   // ---------- 网络 18 ----------
   // 标题：**********************钻孔结束，枪退出速度给定*****************************************
   // 含义：条件 ((((((#DownDrillStep.S20 AND NOT (#DownDrillStep.S22)) AND ("DB720_KuKa_MainCtrl".CmdOut.gi_ToolTypeNo = 2))) AND #DownDrillStep.StopDrill_Ack) AND NOT ("DB1900_Communication_PC".Para.ProduceMode3)) AND ("DB1900_Communication_PC".Para.DrillWidth = 22.0)) 成立时，将 20 传送到 "DB1080_Component".Robot.CTRL_IN.RobotSpeed
   IF ((((((#DownDrillStep.S20 AND NOT (#DownDrillStep.S22)) AND ("DB720_KuKa_MainCtrl".CmdOut.gi_ToolTypeNo = 2))) AND #DownDrillStep.StopDrill_Ack) AND NOT ("DB1900_Communication_PC".Para.ProduceMode3)) AND ("DB1900_Communication_PC".Para.DrillWidth = 22.0)) THEN
       "DB1080_Component".Robot.CTRL_IN.RobotSpeed := 20;
   END_IF;
   // 含义：条件 ((((((#DownDrillStep.S20 AND NOT (#DownDrillStep.S22)) AND ("DB720_KuKa_MainCtrl".CmdOut.gi_ToolTypeNo = 2))) AND #DownDrillStep.StopDrill_Ack) AND NOT ("DB1900_Communication_PC".Para.ProduceMode3)) AND ("DB1900_Communication_PC".Para.DrillWidth = 25.0)) 成立时，将 25 传送到 "DB1080_Component".Robot.CTRL_IN.RobotSpeed
   IF ((((((#DownDrillStep.S20 AND NOT (#DownDrillStep.S22)) AND ("DB720_KuKa_MainCtrl".CmdOut.gi_ToolTypeNo = 2))) AND #DownDrillStep.StopDrill_Ack) AND NOT ("DB1900_Communication_PC".Para.ProduceMode3)) AND ("DB1900_Communication_PC".Para.DrillWidth = 25.0)) THEN
       "DB1080_Component".Robot.CTRL_IN.RobotSpeed := 25;
   END_IF;
   // 含义：条件 ((((((#DownDrillStep.S20 AND NOT (#DownDrillStep.S22)) AND ("DB720_KuKa_MainCtrl".CmdOut.gi_ToolTypeNo = 2))) AND #DownDrillStep.StopDrill_Ack) AND NOT ("DB1900_Communication_PC".Para.ProduceMode3)) AND ("DB1900_Communication_PC".Para.DrillWidth > 25.0)) 成立时，将 30 传送到 "DB1080_Component".Robot.CTRL_IN.RobotSpeed
   IF ((((((#DownDrillStep.S20 AND NOT (#DownDrillStep.S22)) AND ("DB720_KuKa_MainCtrl".CmdOut.gi_ToolTypeNo = 2))) AND #DownDrillStep.StopDrill_Ack) AND NOT ("DB1900_Communication_PC".Para.ProduceMode3)) AND ("DB1900_Communication_PC".Para.DrillWidth > 25.0)) THEN
       "DB1080_Component".Robot.CTRL_IN.RobotSpeed := 30;
   END_IF;
   // 含义：条件 ((((#DownDrillStep.S20 AND NOT (#DownDrillStep.S22)) AND ("DB720_KuKa_MainCtrl".CmdOut.gi_ToolTypeNo = 2))) AND #DownDrillStep.StopDrill_Ack) AND "DB1900_Communication_PC".Para.ProduceMode3 成立时，将 50 传送到 "DB1080_Component".Robot.CTRL_IN.RobotSpeed
   IF ((((#DownDrillStep.S20 AND NOT (#DownDrillStep.S22)) AND ("DB720_KuKa_MainCtrl".CmdOut.gi_ToolTypeNo = 2))) AND #DownDrillStep.StopDrill_Ack) AND "DB1900_Communication_PC".Para.ProduceMode3 THEN
       "DB1080_Component".Robot.CTRL_IN.RobotSpeed := 50;
   END_IF;
   // 含义：条件 ((((((#DownDrillStep.S20 AND NOT (#DownDrillStep.S22)) AND ("DB720_KuKa_MainCtrl".CmdOut.gi_ToolTypeNo = 13))) AND #Aux.StartDrill) AND NOT (#DownDrillStep.StopDrill_Ack)) AND ("DB1900_Communication_PC".Recv.Current_2 > 12.0)) 成立时，将 1 传送到 "DB1080_Component".Robot.CTRL_IN.RobotSpeed
   IF ((((((#DownDrillStep.S20 AND NOT (#DownDrillStep.S22)) AND ("DB720_KuKa_MainCtrl".CmdOut.gi_ToolTypeNo = 13))) AND #Aux.StartDrill) AND NOT (#DownDrillStep.StopDrill_Ack)) AND ("DB1900_Communication_PC".Recv.Current_2 > 12.0)) THEN
       "DB1080_Component".Robot.CTRL_IN.RobotSpeed := 1;
   END_IF;
   // 含义：条件 ((((((#DownDrillStep.S20 AND NOT (#DownDrillStep.S22)) AND ("DB720_KuKa_MainCtrl".CmdOut.gi_ToolTypeNo = 13))) AND #Aux.StartDrill) AND #DownDrillStep.StopDrill_Ack) AND ("DB1900_Communication_PC".Recv.Current_2 < 12.0)) 成立时，将 30 传送到 "DB1080_Component".Robot.CTRL_IN.RobotSpeed
   IF ((((((#DownDrillStep.S20 AND NOT (#DownDrillStep.S22)) AND ("DB720_KuKa_MainCtrl".CmdOut.gi_ToolTypeNo = 13))) AND #Aux.StartDrill) AND #DownDrillStep.StopDrill_Ack) AND ("DB1900_Communication_PC".Recv.Current_2 < 12.0)) THEN
       "DB1080_Component".Robot.CTRL_IN.RobotSpeed := 30;
   END_IF;
   // 含义：条件 ((((((#DownDrillStep.S20 AND NOT (#DownDrillStep.S22)) AND ("DB720_KuKa_MainCtrl".CmdOut.gi_ToolTypeNo = 13))) AND #Aux.StartDrill) AND #DownDrillStep.StopDrill_Ack) AND ("DB1900_Communication_PC".Recv.Current_2 >= 12.0)) 成立时，将 10 传送到 "DB1080_Component".Robot.CTRL_IN.RobotSpeed
   IF ((((((#DownDrillStep.S20 AND NOT (#DownDrillStep.S22)) AND ("DB720_KuKa_MainCtrl".CmdOut.gi_ToolTypeNo = 13))) AND #Aux.StartDrill) AND #DownDrillStep.StopDrill_Ack) AND ("DB1900_Communication_PC".Recv.Current_2 >= 12.0)) THEN
       "DB1080_Component".Robot.CTRL_IN.RobotSpeed := 10;
   END_IF;

   // ---------- 网络 19 ----------
   // 标题：****************故障计数（包含钻超时，低电流，打孔深度超限）**************************
   // 含义：调用计数器实例 "Timer_DownChiselEnd".TON（上升沿计数，当前值写入 CV）
   "Timer_DownChiselEnd".TON(IN := ((((#DownDrillStep.S20 AND NOT (#DownDrillStep.S22)) AND "DB1900_Communication_PC".Para.ProduceMode3) AND "DB720_KuKa_MainCtrl".StatusIn.do_DrilEnd_Pos) AND ("DB1900_Communication_PC".Recv.Current_2 < "DB1900_Communication_PC".Para.CurrentMinLimit)),
                             PT := T#3s);
   // 含义：条件 "Timer_DownChiselEnd".Q 成立时，将 TRUE 传送到 "DB1060_AutoStep".DownDrillAutoStep.DownDrillStep.ChiselEndPos
   IF "Timer_DownChiselEnd".Q THEN
       "DB1060_AutoStep".DownDrillAutoStep.DownDrillStep.ChiselEndPos := TRUE;
   END_IF;
   // 含义：条件 "Timer_DownChiselEnd".Q 成立时，将 ("DB1042_Timer".DCLowTimeOutTimes + 1) 传送到 "DB1042_Timer".DCLowTimeOutTimes
   IF "Timer_DownChiselEnd".Q THEN
       "DB1042_Timer".DCLowTimeOutTimes := ("DB1042_Timer".DCLowTimeOutTimes + 1);
   END_IF;
   // 含义：条件 (((((#DownDrillStep.S20 AND NOT (#DownDrillStep.S22)) AND "DB1900_Communication_PC".Para.ProduceMode3) AND ("DB1900_Communication_PC".Recv.Current_2 > "DB1900_Communication_PC".Para.CurrentMinLimit))) AND ("DB1900_Communication_PC".Recv.Current_2 < "DB1900_Communication_PC".Para.CurrentMaxLimit)) 成立时，将 0 传送到 "DB1042_Timer".DCLowTimeOutTimes
   IF (((((#DownDrillStep.S20 AND NOT (#DownDrillStep.S22)) AND "DB1900_Communication_PC".Para.ProduceMode3) AND ("DB1900_Communication_PC".Recv.Current_2 > "DB1900_Communication_PC".Para.CurrentMinLimit))) AND ("DB1900_Communication_PC".Recv.Current_2 < "DB1900_Communication_PC".Para.CurrentMaxLimit)) THEN
       "DB1042_Timer".DCLowTimeOutTimes := 0;
   END_IF;
   // 含义：条件 ((((#DownDrillStep.S20 AND NOT (#DownDrillStep.S22)) AND "DB1900_Communication_PC".Para.ProduceMode3) AND "DB1042_Timer".DDrillEndTime.Q) OR (((#DownDrillStep.S20 AND NOT (#DownDrillStep.S22)) AND "DB1900_Communication_PC".Para.ProduceMode3) AND #Aux.DDrillTime.Q) OR (((#DownDrillStep.S20 AND NOT (#DownDrillStep.S22)) AND "DB1900_Communication_PC".Para.ProduceMode3) AND "DB1042_Timer".CurrentLowTimeOut.Q) OR (((#DownDrillStep.S20 AND NOT (#DownDrillStep.S22)) AND "DB1900_Communication_PC".Para.ProduceMode3) AND "DB1042_Timer".CurrentHighTimeOut.Q) OR (((#DownDrillStep.S20 AND NOT (#DownDrillStep.S22)) AND "DB1900_Communication_PC".Para.ProduceMode3) AND "DB1060_AutoStep".DownDrillAutoStep.DownDrillStep.ChiselEndPos) OR ((((#DownDrillStep.S20 AND NOT (#DownDrillStep.S22)) AND "DB1900_Communication_PC".Para.ProduceMode3) AND ("DB1900_Communication_PC".Send.ScrLen >= "DB1900_Communication_PC".Para.DrillDepth)))) AND NOT ("DB720_KuKa_MainCtrl".StatusIn.do_ChiselCylinderExt) 成立时，将 0.0 传送到 "DB1080_Component".Aux.Pressure
   IF ((((#DownDrillStep.S20 AND NOT (#DownDrillStep.S22)) AND "DB1900_Communication_PC".Para.ProduceMode3) AND "DB1042_Timer".DDrillEndTime.Q) OR (((#DownDrillStep.S20 AND NOT (#DownDrillStep.S22)) AND "DB1900_Communication_PC".Para.ProduceMode3) AND #Aux.DDrillTime.Q) OR (((#DownDrillStep.S20 AND NOT (#DownDrillStep.S22)) AND "DB1900_Communication_PC".Para.ProduceMode3) AND "DB1042_Timer".CurrentLowTimeOut.Q) OR (((#DownDrillStep.S20 AND NOT (#DownDrillStep.S22)) AND "DB1900_Communication_PC".Para.ProduceMode3) AND "DB1042_Timer".CurrentHighTimeOut.Q) OR (((#DownDrillStep.S20 AND NOT (#DownDrillStep.S22)) AND "DB1900_Communication_PC".Para.ProduceMode3) AND "DB1060_AutoStep".DownDrillAutoStep.DownDrillStep.ChiselEndPos) OR ((((#DownDrillStep.S20 AND NOT (#DownDrillStep.S22)) AND "DB1900_Communication_PC".Para.ProduceMode3) AND ("DB1900_Communication_PC".Send.ScrLen >= "DB1900_Communication_PC".Para.DrillDepth)))) AND NOT ("DB720_KuKa_MainCtrl".StatusIn.do_ChiselCylinderExt) THEN
       "DB1080_Component".Aux.Pressure := 0.0;
   END_IF;
   // 含义：条件 ((((#DownDrillStep.S20 AND NOT (#DownDrillStep.S22)) AND "DB1900_Communication_PC".Para.ProduceMode3) AND "DB1042_Timer".DDrillEndTime.Q) OR (((#DownDrillStep.S20 AND NOT (#DownDrillStep.S22)) AND "DB1900_Communication_PC".Para.ProduceMode3) AND #Aux.DDrillTime.Q) OR (((#DownDrillStep.S20 AND NOT (#DownDrillStep.S22)) AND "DB1900_Communication_PC".Para.ProduceMode3) AND "DB1042_Timer".CurrentLowTimeOut.Q) OR (((#DownDrillStep.S20 AND NOT (#DownDrillStep.S22)) AND "DB1900_Communication_PC".Para.ProduceMode3) AND "DB1042_Timer".CurrentHighTimeOut.Q) OR (((#DownDrillStep.S20 AND NOT (#DownDrillStep.S22)) AND "DB1900_Communication_PC".Para.ProduceMode3) AND "DB1060_AutoStep".DownDrillAutoStep.DownDrillStep.ChiselEndPos) OR ((((#DownDrillStep.S20 AND NOT (#DownDrillStep.S22)) AND "DB1900_Communication_PC".Para.ProduceMode3) AND ("DB1900_Communication_PC".Send.ScrLen >= "DB1900_Communication_PC".Para.DrillDepth)))) AND NOT ("DB720_KuKa_MainCtrl".CmdOut.di_ChiselRobotRet) 成立时，将 TRUE 传送到 "DB1081_ValveCall".ST01.Z02.RetAuto
   IF ((((#DownDrillStep.S20 AND NOT (#DownDrillStep.S22)) AND "DB1900_Communication_PC".Para.ProduceMode3) AND "DB1042_Timer".DDrillEndTime.Q) OR (((#DownDrillStep.S20 AND NOT (#DownDrillStep.S22)) AND "DB1900_Communication_PC".Para.ProduceMode3) AND #Aux.DDrillTime.Q) OR (((#DownDrillStep.S20 AND NOT (#DownDrillStep.S22)) AND "DB1900_Communication_PC".Para.ProduceMode3) AND "DB1042_Timer".CurrentLowTimeOut.Q) OR (((#DownDrillStep.S20 AND NOT (#DownDrillStep.S22)) AND "DB1900_Communication_PC".Para.ProduceMode3) AND "DB1042_Timer".CurrentHighTimeOut.Q) OR (((#DownDrillStep.S20 AND NOT (#DownDrillStep.S22)) AND "DB1900_Communication_PC".Para.ProduceMode3) AND "DB1060_AutoStep".DownDrillAutoStep.DownDrillStep.ChiselEndPos) OR ((((#DownDrillStep.S20 AND NOT (#DownDrillStep.S22)) AND "DB1900_Communication_PC".Para.ProduceMode3) AND ("DB1900_Communication_PC".Send.ScrLen >= "DB1900_Communication_PC".Para.DrillDepth)))) AND NOT ("DB720_KuKa_MainCtrl".CmdOut.di_ChiselRobotRet) THEN
       "DB1081_ValveCall".ST01.Z02.RetAuto := TRUE;
   END_IF;
   // 含义：条件 ((((#DownDrillStep.S20 AND NOT (#DownDrillStep.S22)) AND "DB1900_Communication_PC".Para.ProduceMode3) AND "DB1042_Timer".DDrillEndTime.Q) OR (((#DownDrillStep.S20 AND NOT (#DownDrillStep.S22)) AND "DB1900_Communication_PC".Para.ProduceMode3) AND #Aux.DDrillTime.Q) OR (((#DownDrillStep.S20 AND NOT (#DownDrillStep.S22)) AND "DB1900_Communication_PC".Para.ProduceMode3) AND "DB1042_Timer".CurrentLowTimeOut.Q) OR (((#DownDrillStep.S20 AND NOT (#DownDrillStep.S22)) AND "DB1900_Communication_PC".Para.ProduceMode3) AND "DB1042_Timer".CurrentHighTimeOut.Q) OR (((#DownDrillStep.S20 AND NOT (#DownDrillStep.S22)) AND "DB1900_Communication_PC".Para.ProduceMode3) AND "DB1060_AutoStep".DownDrillAutoStep.DownDrillStep.ChiselEndPos) OR ((((#DownDrillStep.S20 AND NOT (#DownDrillStep.S22)) AND "DB1900_Communication_PC".Para.ProduceMode3) AND ("DB1900_Communication_PC".Send.ScrLen >= "DB1900_Communication_PC".Para.DrillDepth)))) AND "DB720_KuKa_MainCtrl".StatusIn.do_ChiselCylinderExt 成立时，将 FALSE 传送到 "DB1081_ValveCall".ST01.Z02.RetAuto
   IF ((((#DownDrillStep.S20 AND NOT (#DownDrillStep.S22)) AND "DB1900_Communication_PC".Para.ProduceMode3) AND "DB1042_Timer".DDrillEndTime.Q) OR (((#DownDrillStep.S20 AND NOT (#DownDrillStep.S22)) AND "DB1900_Communication_PC".Para.ProduceMode3) AND #Aux.DDrillTime.Q) OR (((#DownDrillStep.S20 AND NOT (#DownDrillStep.S22)) AND "DB1900_Communication_PC".Para.ProduceMode3) AND "DB1042_Timer".CurrentLowTimeOut.Q) OR (((#DownDrillStep.S20 AND NOT (#DownDrillStep.S22)) AND "DB1900_Communication_PC".Para.ProduceMode3) AND "DB1042_Timer".CurrentHighTimeOut.Q) OR (((#DownDrillStep.S20 AND NOT (#DownDrillStep.S22)) AND "DB1900_Communication_PC".Para.ProduceMode3) AND "DB1060_AutoStep".DownDrillAutoStep.DownDrillStep.ChiselEndPos) OR ((((#DownDrillStep.S20 AND NOT (#DownDrillStep.S22)) AND "DB1900_Communication_PC".Para.ProduceMode3) AND ("DB1900_Communication_PC".Send.ScrLen >= "DB1900_Communication_PC".Para.DrillDepth)))) AND "DB720_KuKa_MainCtrl".StatusIn.do_ChiselCylinderExt THEN
       "DB1081_ValveCall".ST01.Z02.RetAuto := FALSE;
   END_IF;
   // 含义：条件 ((((#DownDrillStep.S20 AND NOT (#DownDrillStep.S22)) AND "DB1900_Communication_PC".Para.ProduceMode3) AND "DB1042_Timer".DDrillEndTime.Q) OR (((#DownDrillStep.S20 AND NOT (#DownDrillStep.S22)) AND "DB1900_Communication_PC".Para.ProduceMode3) AND #Aux.DDrillTime.Q) OR (((#DownDrillStep.S20 AND NOT (#DownDrillStep.S22)) AND "DB1900_Communication_PC".Para.ProduceMode3) AND "DB1042_Timer".CurrentLowTimeOut.Q) OR (((#DownDrillStep.S20 AND NOT (#DownDrillStep.S22)) AND "DB1900_Communication_PC".Para.ProduceMode3) AND "DB1042_Timer".CurrentHighTimeOut.Q) OR (((#DownDrillStep.S20 AND NOT (#DownDrillStep.S22)) AND "DB1900_Communication_PC".Para.ProduceMode3) AND "DB1060_AutoStep".DownDrillAutoStep.DownDrillStep.ChiselEndPos) OR ((((#DownDrillStep.S20 AND NOT (#DownDrillStep.S22)) AND "DB1900_Communication_PC".Para.ProduceMode3) AND ("DB1900_Communication_PC".Send.ScrLen >= "DB1900_Communication_PC".Para.DrillDepth)))) AND "DB720_KuKa_MainCtrl".StatusIn.do_ReqStopDril 成立时，将 FALSE 传送到 "DB720_KuKa_MainCtrl".CmdOut.di_ChiselCylinderRet
   IF ((((#DownDrillStep.S20 AND NOT (#DownDrillStep.S22)) AND "DB1900_Communication_PC".Para.ProduceMode3) AND "DB1042_Timer".DDrillEndTime.Q) OR (((#DownDrillStep.S20 AND NOT (#DownDrillStep.S22)) AND "DB1900_Communication_PC".Para.ProduceMode3) AND #Aux.DDrillTime.Q) OR (((#DownDrillStep.S20 AND NOT (#DownDrillStep.S22)) AND "DB1900_Communication_PC".Para.ProduceMode3) AND "DB1042_Timer".CurrentLowTimeOut.Q) OR (((#DownDrillStep.S20 AND NOT (#DownDrillStep.S22)) AND "DB1900_Communication_PC".Para.ProduceMode3) AND "DB1042_Timer".CurrentHighTimeOut.Q) OR (((#DownDrillStep.S20 AND NOT (#DownDrillStep.S22)) AND "DB1900_Communication_PC".Para.ProduceMode3) AND "DB1060_AutoStep".DownDrillAutoStep.DownDrillStep.ChiselEndPos) OR ((((#DownDrillStep.S20 AND NOT (#DownDrillStep.S22)) AND "DB1900_Communication_PC".Para.ProduceMode3) AND ("DB1900_Communication_PC".Send.ScrLen >= "DB1900_Communication_PC".Para.DrillDepth)))) AND "DB720_KuKa_MainCtrl".StatusIn.do_ReqStopDril THEN
       "DB720_KuKa_MainCtrl".CmdOut.di_ChiselCylinderRet := FALSE;
   END_IF;
   // 含义：条件 ((((#DownDrillStep.S20 AND NOT (#DownDrillStep.S22)) AND "DB1900_Communication_PC".Para.ProduceMode3) AND "DB1042_Timer".DDrillEndTime.Q) OR (((#DownDrillStep.S20 AND NOT (#DownDrillStep.S22)) AND "DB1900_Communication_PC".Para.ProduceMode3) AND #Aux.DDrillTime.Q) OR (((#DownDrillStep.S20 AND NOT (#DownDrillStep.S22)) AND "DB1900_Communication_PC".Para.ProduceMode3) AND "DB1042_Timer".CurrentLowTimeOut.Q) OR (((#DownDrillStep.S20 AND NOT (#DownDrillStep.S22)) AND "DB1900_Communication_PC".Para.ProduceMode3) AND "DB1042_Timer".CurrentHighTimeOut.Q) OR (((#DownDrillStep.S20 AND NOT (#DownDrillStep.S22)) AND "DB1900_Communication_PC".Para.ProduceMode3) AND "DB1060_AutoStep".DownDrillAutoStep.DownDrillStep.ChiselEndPos) OR ((((#DownDrillStep.S20 AND NOT (#DownDrillStep.S22)) AND "DB1900_Communication_PC".Para.ProduceMode3) AND ("DB1900_Communication_PC".Send.ScrLen >= "DB1900_Communication_PC".Para.DrillDepth)))) AND "DB720_KuKa_MainCtrl".StatusIn.do_ReqStopDril 成立时，将 FALSE 传送到 "DB720_KuKa_MainCtrl".CmdOut.di_ChiselRobotRet
   IF ((((#DownDrillStep.S20 AND NOT (#DownDrillStep.S22)) AND "DB1900_Communication_PC".Para.ProduceMode3) AND "DB1042_Timer".DDrillEndTime.Q) OR (((#DownDrillStep.S20 AND NOT (#DownDrillStep.S22)) AND "DB1900_Communication_PC".Para.ProduceMode3) AND #Aux.DDrillTime.Q) OR (((#DownDrillStep.S20 AND NOT (#DownDrillStep.S22)) AND "DB1900_Communication_PC".Para.ProduceMode3) AND "DB1042_Timer".CurrentLowTimeOut.Q) OR (((#DownDrillStep.S20 AND NOT (#DownDrillStep.S22)) AND "DB1900_Communication_PC".Para.ProduceMode3) AND "DB1042_Timer".CurrentHighTimeOut.Q) OR (((#DownDrillStep.S20 AND NOT (#DownDrillStep.S22)) AND "DB1900_Communication_PC".Para.ProduceMode3) AND "DB1060_AutoStep".DownDrillAutoStep.DownDrillStep.ChiselEndPos) OR ((((#DownDrillStep.S20 AND NOT (#DownDrillStep.S22)) AND "DB1900_Communication_PC".Para.ProduceMode3) AND ("DB1900_Communication_PC".Send.ScrLen >= "DB1900_Communication_PC".Para.DrillDepth)))) AND "DB720_KuKa_MainCtrl".StatusIn.do_ReqStopDril THEN
       "DB720_KuKa_MainCtrl".CmdOut.di_ChiselRobotRet := FALSE;
   END_IF;
   // 含义：条件 ((((((#DownDrillStep.S20 AND NOT (#DownDrillStep.S22)) AND "DB1900_Communication_PC".Para.ProduceMode3) AND "DB1042_Timer".DDrillEndTime.Q) OR (((#DownDrillStep.S20 AND NOT (#DownDrillStep.S22)) AND "DB1900_Communication_PC".Para.ProduceMode3) AND #Aux.DDrillTime.Q) OR (((#DownDrillStep.S20 AND NOT (#DownDrillStep.S22)) AND "DB1900_Communication_PC".Para.ProduceMode3) AND "DB1042_Timer".CurrentLowTimeOut.Q) OR (((#DownDrillStep.S20 AND NOT (#DownDrillStep.S22)) AND "DB1900_Communication_PC".Para.ProduceMode3) AND "DB1042_Timer".CurrentHighTimeOut.Q) OR (((#DownDrillStep.S20 AND NOT (#DownDrillStep.S22)) AND "DB1900_Communication_PC".Para.ProduceMode3) AND "DB1060_AutoStep".DownDrillAutoStep.DownDrillStep.ChiselEndPos) OR ((((#DownDrillStep.S20 AND NOT (#DownDrillStep.S22)) AND "DB1900_Communication_PC".Para.ProduceMode3) AND ("DB1900_Communication_PC".Send.ScrLen >= "DB1900_Communication_PC".Para.DrillDepth)))) AND "IZ02RetPos") AND ("DB1080_Component".ClinyderPos.Ctrl_Out.Cur_Val_Out >= 92.5)) 成立时，将 TRUE 传送到 "DB720_KuKa_MainCtrl".CmdOut.di_ChiselCylinderRet
   IF ((((((#DownDrillStep.S20 AND NOT (#DownDrillStep.S22)) AND "DB1900_Communication_PC".Para.ProduceMode3) AND "DB1042_Timer".DDrillEndTime.Q) OR (((#DownDrillStep.S20 AND NOT (#DownDrillStep.S22)) AND "DB1900_Communication_PC".Para.ProduceMode3) AND #Aux.DDrillTime.Q) OR (((#DownDrillStep.S20 AND NOT (#DownDrillStep.S22)) AND "DB1900_Communication_PC".Para.ProduceMode3) AND "DB1042_Timer".CurrentLowTimeOut.Q) OR (((#DownDrillStep.S20 AND NOT (#DownDrillStep.S22)) AND "DB1900_Communication_PC".Para.ProduceMode3) AND "DB1042_Timer".CurrentHighTimeOut.Q) OR (((#DownDrillStep.S20 AND NOT (#DownDrillStep.S22)) AND "DB1900_Communication_PC".Para.ProduceMode3) AND "DB1060_AutoStep".DownDrillAutoStep.DownDrillStep.ChiselEndPos) OR ((((#DownDrillStep.S20 AND NOT (#DownDrillStep.S22)) AND "DB1900_Communication_PC".Para.ProduceMode3) AND ("DB1900_Communication_PC".Send.ScrLen >= "DB1900_Communication_PC".Para.DrillDepth)))) AND "IZ02RetPos") AND ("DB1080_Component".ClinyderPos.Ctrl_Out.Cur_Val_Out >= 92.5)) THEN
       "DB720_KuKa_MainCtrl".CmdOut.di_ChiselCylinderRet := TRUE;
   END_IF;
   // 含义：条件 ((((((#DownDrillStep.S20 AND NOT (#DownDrillStep.S22)) AND "DB1900_Communication_PC".Para.ProduceMode3) AND "DB1042_Timer".DDrillEndTime.Q) OR (((#DownDrillStep.S20 AND NOT (#DownDrillStep.S22)) AND "DB1900_Communication_PC".Para.ProduceMode3) AND #Aux.DDrillTime.Q) OR (((#DownDrillStep.S20 AND NOT (#DownDrillStep.S22)) AND "DB1900_Communication_PC".Para.ProduceMode3) AND "DB1042_Timer".CurrentLowTimeOut.Q) OR (((#DownDrillStep.S20 AND NOT (#DownDrillStep.S22)) AND "DB1900_Communication_PC".Para.ProduceMode3) AND "DB1042_Timer".CurrentHighTimeOut.Q) OR (((#DownDrillStep.S20 AND NOT (#DownDrillStep.S22)) AND "DB1900_Communication_PC".Para.ProduceMode3) AND "DB1060_AutoStep".DownDrillAutoStep.DownDrillStep.ChiselEndPos) OR ((((#DownDrillStep.S20 AND NOT (#DownDrillStep.S22)) AND "DB1900_Communication_PC".Para.ProduceMode3) AND ("DB1900_Communication_PC".Send.ScrLen >= "DB1900_Communication_PC".Para.DrillDepth)))) AND "IZ02RetPos") AND ("DB1080_Component".ClinyderPos.Ctrl_Out.Cur_Val_Out >= 92.5)) 成立时，将 TRUE 传送到 "DB720_KuKa_MainCtrl".CmdOut.di_ChiselRobotRet
   IF ((((((#DownDrillStep.S20 AND NOT (#DownDrillStep.S22)) AND "DB1900_Communication_PC".Para.ProduceMode3) AND "DB1042_Timer".DDrillEndTime.Q) OR (((#DownDrillStep.S20 AND NOT (#DownDrillStep.S22)) AND "DB1900_Communication_PC".Para.ProduceMode3) AND #Aux.DDrillTime.Q) OR (((#DownDrillStep.S20 AND NOT (#DownDrillStep.S22)) AND "DB1900_Communication_PC".Para.ProduceMode3) AND "DB1042_Timer".CurrentLowTimeOut.Q) OR (((#DownDrillStep.S20 AND NOT (#DownDrillStep.S22)) AND "DB1900_Communication_PC".Para.ProduceMode3) AND "DB1042_Timer".CurrentHighTimeOut.Q) OR (((#DownDrillStep.S20 AND NOT (#DownDrillStep.S22)) AND "DB1900_Communication_PC".Para.ProduceMode3) AND "DB1060_AutoStep".DownDrillAutoStep.DownDrillStep.ChiselEndPos) OR ((((#DownDrillStep.S20 AND NOT (#DownDrillStep.S22)) AND "DB1900_Communication_PC".Para.ProduceMode3) AND ("DB1900_Communication_PC".Send.ScrLen >= "DB1900_Communication_PC".Para.DrillDepth)))) AND "IZ02RetPos") AND ("DB1080_Component".ClinyderPos.Ctrl_Out.Cur_Val_Out >= 92.5)) THEN
       "DB720_KuKa_MainCtrl".CmdOut.di_ChiselRobotRet := TRUE;
   END_IF;
   // 含义：调用计数器实例 "Timer_CylinderBack_Down".TON（上升沿计数，当前值写入 CV）
   "Timer_CylinderBack_Down".TON(IN := ((((#DownDrillStep.S20 AND NOT (#DownDrillStep.S22)) AND "DB1900_Communication_PC".Para.ProduceMode3) AND "DB1042_Timer".DDrillEndTime.Q) OR (((#DownDrillStep.S20 AND NOT (#DownDrillStep.S22)) AND "DB1900_Communication_PC".Para.ProduceMode3) AND #Aux.DDrillTime.Q) OR (((#DownDrillStep.S20 AND NOT (#DownDrillStep.S22)) AND "DB1900_Communication_PC".Para.ProduceMode3) AND "DB1042_Timer".CurrentLowTimeOut.Q) OR (((#DownDrillStep.S20 AND NOT (#DownDrillStep.S22)) AND "DB1900_Communication_PC".Para.ProduceMode3) AND "DB1042_Timer".CurrentHighTimeOut.Q) OR (((#DownDrillStep.S20 AND NOT (#DownDrillStep.S22)) AND "DB1900_Communication_PC".Para.ProduceMode3) AND "DB1060_AutoStep".DownDrillAutoStep.DownDrillStep.ChiselEndPos) OR ((((#DownDrillStep.S20 AND NOT (#DownDrillStep.S22)) AND "DB1900_Communication_PC".Para.ProduceMode3) AND ("DB1900_Communication_PC".Send.ScrLen >= "DB1900_Communication_PC".Para.DrillDepth)))) AND NOT ("IZ02RetPos"),
                                 PT := t#3s);
   // 含义：条件 "Timer_CylinderBack_Down".Q 成立时，将 TRUE 传送到 "DB720_KuKa_MainCtrl".CmdOut.di_ChiselRobotRet
   IF "Timer_CylinderBack_Down".Q THEN
       "DB720_KuKa_MainCtrl".CmdOut.di_ChiselRobotRet := TRUE;
   END_IF;
   // 含义：调用计数器实例 "Timer_RobotPry_Down".TON（上升沿计数，当前值写入 CV）
   "Timer_RobotPry_Down".TON(IN := (((((#DownDrillStep.S20 AND NOT (#DownDrillStep.S22)) AND "DB1900_Communication_PC".Para.ProduceMode3) AND "DB1042_Timer".DDrillEndTime.Q) OR (((#DownDrillStep.S20 AND NOT (#DownDrillStep.S22)) AND "DB1900_Communication_PC".Para.ProduceMode3) AND #Aux.DDrillTime.Q) OR (((#DownDrillStep.S20 AND NOT (#DownDrillStep.S22)) AND "DB1900_Communication_PC".Para.ProduceMode3) AND "DB1042_Timer".CurrentLowTimeOut.Q) OR (((#DownDrillStep.S20 AND NOT (#DownDrillStep.S22)) AND "DB1900_Communication_PC".Para.ProduceMode3) AND "DB1042_Timer".CurrentHighTimeOut.Q) OR (((#DownDrillStep.S20 AND NOT (#DownDrillStep.S22)) AND "DB1900_Communication_PC".Para.ProduceMode3) AND "DB1060_AutoStep".DownDrillAutoStep.DownDrillStep.ChiselEndPos) OR ((((#DownDrillStep.S20 AND NOT (#DownDrillStep.S22)) AND "DB1900_Communication_PC".Para.ProduceMode3) AND ("DB1900_Communication_PC".Send.ScrLen >= "DB1900_Communication_PC".Para.DrillDepth)))) AND NOT ("IZ02RetPos")) AND "DB720_KuKa_MainCtrl".StatusIn.do_RobotPry_End,
                             PT := t#3s);
   // 含义：条件 "Timer_RobotPry_Down".Q 成立时，将 FALSE 传送到 "DB720_KuKa_MainCtrl".CmdOut.di_ChiselCylinderRet
   IF "Timer_RobotPry_Down".Q THEN
       "DB720_KuKa_MainCtrl".CmdOut.di_ChiselCylinderRet := FALSE;
   END_IF;
   // 含义：条件 "Timer_RobotPry_Down".Q 成立时，将 FALSE 传送到 "DB720_KuKa_MainCtrl".CmdOut.di_ChiselRobotRet
   IF "Timer_RobotPry_Down".Q THEN
       "DB720_KuKa_MainCtrl".CmdOut.di_ChiselRobotRet := FALSE;
   END_IF;
   // 含义：条件 "Timer_RobotPry_Down".Q 成立时，将 TRUE 传送到 "DB1148_PromptBeeper".Public.DownChiselStuckErr
   IF "Timer_RobotPry_Down".Q THEN
       "DB1148_PromptBeeper".Public.DownChiselStuckErr := TRUE;
   END_IF;
   // 含义：条件 "Timer_RobotPry_Down".Q 成立时，将 TRUE 传送到 #DownDrillStep.ErrEnd
   IF "Timer_RobotPry_Down".Q THEN
       #DownDrillStep.ErrEnd := TRUE;
   END_IF;
   // 含义：条件 "Timer_RobotPry_Down".Q 成立时，将 FALSE 传送到 "DB1081_ValveCall".ST01.Z02.RetAuto
   IF "Timer_RobotPry_Down".Q THEN
       "DB1081_ValveCall".ST01.Z02.RetAuto := FALSE;
   END_IF;
   // 含义：条件 "Timer_RobotPry_Down".Q 成立时，将 TRUE 传送到 "DB1081_ValveCall".ST01.Z01.ExtAuto
   IF "Timer_RobotPry_Down".Q THEN
       "DB1081_ValveCall".ST01.Z01.ExtAuto := TRUE;
   END_IF;
   // 含义：条件 "Timer_RobotPry_Down".Q 成立时，将 FALSE 传送到 "DB1081_ValveCall".ST01.Z01.RetAuto
   IF "Timer_RobotPry_Down".Q THEN
       "DB1081_ValveCall".ST01.Z01.RetAuto := FALSE;
   END_IF;
   // 含义：条件 "Timer_RobotPry_Down".Q 成立时，将 0.1 传送到 "DB1080_Component".Aux.Pressure
   IF "Timer_RobotPry_Down".Q THEN
       "DB1080_Component".Aux.Pressure := 0.1;
   END_IF;
   // 含义：将 (((#DownDrillStep.S20 AND NOT (#DownDrillStep.S22)) AND #Aux.DDrillTime.Q) OR ((#DownDrillStep.S20 AND NOT (#DownDrillStep.S22)) AND "DB1042_Timer".CurrentLowTimeOut.Q) OR ((#DownDrillStep.S20 AND NOT (#DownDrillStep.S22)) AND "DB1042_Timer".CurrentHighTimeOut.Q) OR ((((((((#DownDrillStep.S20 AND NOT (#DownDrillStep.S22)) AND NOT ("DB1900_Communication_PC".Para.ProduceMode3)) AND ("DB1900_Communication_PC".Send.PosNo <= 2))) AND ("DB1900_Communication_PC".Para.DrillWidth <= 28.0))) AND ("DB1900_Communication_PC".Send.ScrLen >= 55.0))) OR ((((#DownDrillStep.S20 AND NOT (#DownDrillStep.S22)) AND NOT ("DB1900_Communication_PC".Para.ProduceMode3)) AND ("DB1900_Communication_PC".Send.ScrLen >= "DB1900_Communication_PC".Para.DrillDepth))) OR (((#DownDrillStep.S20 AND NOT (#DownDrillStep.S22)) AND "DB1042_Timer".DDrillEndTime.Q) AND "DB1900_Communication_PC".Para.DrillEndMode)) AND NOT ("DB1900_Communication_PC".Para.ProduceMode3) 赋给 #DownDrillStep.StopDrill_End
   #DownDrillStep.StopDrill_End := (((#DownDrillStep.S20 AND NOT (#DownDrillStep.S22)) AND #Aux.DDrillTime.Q) OR ((#DownDrillStep.S20 AND NOT (#DownDrillStep.S22)) AND "DB1042_Timer".CurrentLowTimeOut.Q) OR ((#DownDrillStep.S20 AND NOT (#DownDrillStep.S22)) AND "DB1042_Timer".CurrentHighTimeOut.Q) OR ((((((((#DownDrillStep.S20 AND NOT (#DownDrillStep.S22)) AND NOT ("DB1900_Communication_PC".Para.ProduceMode3)) AND ("DB1900_Communication_PC".Send.PosNo <= 2))) AND ("DB1900_Communication_PC".Para.DrillWidth <= 28.0))) AND ("DB1900_Communication_PC".Send.ScrLen >= 55.0))) OR ((((#DownDrillStep.S20 AND NOT (#DownDrillStep.S22)) AND NOT ("DB1900_Communication_PC".Para.ProduceMode3)) AND ("DB1900_Communication_PC".Send.ScrLen >= "DB1900_Communication_PC".Para.DrillDepth))) OR (((#DownDrillStep.S20 AND NOT (#DownDrillStep.S22)) AND "DB1042_Timer".DDrillEndTime.Q) AND "DB1900_Communication_PC".Para.DrillEndMode)) AND NOT ("DB1900_Communication_PC".Para.ProduceMode3);
   // 含义：条件 ((#DownDrillStep.S20 AND NOT (#DownDrillStep.S22)) AND TRUE) AND "DB1042_Timer".CurrentLowTimeOut.Q 成立时，将 ("DB1042_Timer".DCLowTimeOutTimes + 1) 传送到 "DB1042_Timer".DCLowTimeOutTimes
   IF ((#DownDrillStep.S20 AND NOT (#DownDrillStep.S22)) AND TRUE) AND "DB1042_Timer".CurrentLowTimeOut.Q THEN
       "DB1042_Timer".DCLowTimeOutTimes := ("DB1042_Timer".DCLowTimeOutTimes + 1);
   END_IF;
   // 含义：条件 ((#DownDrillStep.S20 AND NOT (#DownDrillStep.S22)) AND TRUE) AND "DB1042_Timer".CurrentHighTimeOut.Q 成立时，将 ("DB1042_Timer".DCHighTimeOutTimes + 1) 传送到 "DB1042_Timer".DCHighTimeOutTimes
   IF ((#DownDrillStep.S20 AND NOT (#DownDrillStep.S22)) AND TRUE) AND "DB1042_Timer".CurrentHighTimeOut.Q THEN
       "DB1042_Timer".DCHighTimeOutTimes := ("DB1042_Timer".DCHighTimeOutTimes + 1);
   END_IF;
   // 含义：条件 ((((#DownDrillStep.S20 AND NOT (#DownDrillStep.S22)) AND TRUE) AND #Aux.DDrillTime.Q) AND NOT ("DB1900_Communication_PC".Para.DrillEndMode)) OR (((((#DownDrillStep.S20 AND NOT (#DownDrillStep.S22)) AND TRUE) AND #Aux.DDrillTime.Q) AND "DB1900_Communication_PC".Para.ProduceMode3) AND "DB1900_Communication_PC".Para.DrillEndMode) 成立时，将 ("DB1042_Timer".DTimeOutTimes + 1) 传送到 "DB1042_Timer".DTimeOutTimes
   IF ((((#DownDrillStep.S20 AND NOT (#DownDrillStep.S22)) AND TRUE) AND #Aux.DDrillTime.Q) AND NOT ("DB1900_Communication_PC".Para.DrillEndMode)) OR (((((#DownDrillStep.S20 AND NOT (#DownDrillStep.S22)) AND TRUE) AND #Aux.DDrillTime.Q) AND "DB1900_Communication_PC".Para.ProduceMode3) AND "DB1900_Communication_PC".Para.DrillEndMode) THEN
       "DB1042_Timer".DTimeOutTimes := ("DB1042_Timer".DTimeOutTimes + 1);
   END_IF;
   // 含义：条件 (((#DownDrillStep.S20 AND NOT (#DownDrillStep.S22)) AND TRUE) AND ("DB1042_Timer".DCLowTimeOutTimes > 2)) 成立时，将 TRUE 传送到 "DB1148_PromptBeeper".Public.CurrentLowTimeOut
   IF (((#DownDrillStep.S20 AND NOT (#DownDrillStep.S22)) AND TRUE) AND ("DB1042_Timer".DCLowTimeOutTimes > 2)) THEN
       "DB1148_PromptBeeper".Public.CurrentLowTimeOut := TRUE;
   END_IF;
   // 含义：条件 (((#DownDrillStep.S20 AND NOT (#DownDrillStep.S22)) AND TRUE) AND ("DB1042_Timer".DCLowTimeOutTimes > 2)) 成立时，将 TRUE 传送到 #DownDrillStep.ErrEnd
   IF (((#DownDrillStep.S20 AND NOT (#DownDrillStep.S22)) AND TRUE) AND ("DB1042_Timer".DCLowTimeOutTimes > 2)) THEN
       #DownDrillStep.ErrEnd := TRUE;
   END_IF;
   // 含义：条件 (((#DownDrillStep.S20 AND NOT (#DownDrillStep.S22)) AND TRUE) AND ("DB1042_Timer".DCLowTimeOutTimes > 2)) 成立时，将 0 传送到 "DB1042_Timer".DCLowTimeOutTimes
   IF (((#DownDrillStep.S20 AND NOT (#DownDrillStep.S22)) AND TRUE) AND ("DB1042_Timer".DCLowTimeOutTimes > 2)) THEN
       "DB1042_Timer".DCLowTimeOutTimes := 0;
   END_IF;
   // 含义：条件 (((#DownDrillStep.S20 AND NOT (#DownDrillStep.S22)) AND TRUE) AND ("DB1042_Timer".DCHighTimeOutTimes > 2)) 成立时，将 TRUE 传送到 "DB1148_PromptBeeper".Public.CurrentHighTimeOut
   IF (((#DownDrillStep.S20 AND NOT (#DownDrillStep.S22)) AND TRUE) AND ("DB1042_Timer".DCHighTimeOutTimes > 2)) THEN
       "DB1148_PromptBeeper".Public.CurrentHighTimeOut := TRUE;
   END_IF;
   // 含义：条件 (((#DownDrillStep.S20 AND NOT (#DownDrillStep.S22)) AND TRUE) AND ("DB1042_Timer".DCHighTimeOutTimes > 2)) 成立时，将 TRUE 传送到 #DownDrillStep.ErrEnd
   IF (((#DownDrillStep.S20 AND NOT (#DownDrillStep.S22)) AND TRUE) AND ("DB1042_Timer".DCHighTimeOutTimes > 2)) THEN
       #DownDrillStep.ErrEnd := TRUE;
   END_IF;
   // 含义：条件 (((#DownDrillStep.S20 AND NOT (#DownDrillStep.S22)) AND TRUE) AND ("DB1042_Timer".DCHighTimeOutTimes > 2)) 成立时，将 0 传送到 "DB1042_Timer".DCHighTimeOutTimes
   IF (((#DownDrillStep.S20 AND NOT (#DownDrillStep.S22)) AND TRUE) AND ("DB1042_Timer".DCHighTimeOutTimes > 2)) THEN
       "DB1042_Timer".DCHighTimeOutTimes := 0;
   END_IF;
   // 含义：条件 (((#DownDrillStep.S20 AND NOT (#DownDrillStep.S22)) AND TRUE) AND ("DB1042_Timer".DTimeOutTimes > 2)) 成立时，将 TRUE 传送到 #DownDrillStep.ErrEnd
   IF (((#DownDrillStep.S20 AND NOT (#DownDrillStep.S22)) AND TRUE) AND ("DB1042_Timer".DTimeOutTimes > 2)) THEN
       #DownDrillStep.ErrEnd := TRUE;
   END_IF;
   // 含义：条件 (((#DownDrillStep.S20 AND NOT (#DownDrillStep.S22)) AND TRUE) AND ("DB1042_Timer".DTimeOutTimes > 2)) 成立时，将 TRUE 传送到 "DB1148_PromptBeeper".Public.DrillTimeOut
   IF (((#DownDrillStep.S20 AND NOT (#DownDrillStep.S22)) AND TRUE) AND ("DB1042_Timer".DTimeOutTimes > 2)) THEN
       "DB1148_PromptBeeper".Public.DrillTimeOut := TRUE;
   END_IF;
   // 含义：条件 (((#DownDrillStep.S20 AND NOT (#DownDrillStep.S22)) AND TRUE) AND ("DB1042_Timer".DTimeOutTimes > 2)) 成立时，将 0 传送到 "DB1042_Timer".DTimeOutTimes
   IF (((#DownDrillStep.S20 AND NOT (#DownDrillStep.S22)) AND TRUE) AND ("DB1042_Timer".DTimeOutTimes > 2)) THEN
       "DB1042_Timer".DTimeOutTimes := 0;
   END_IF;
   // 含义：条件 (((#DownDrillStep.S20 AND NOT (#DownDrillStep.S22)) AND TRUE) AND ("DB1900_Communication_PC".Send.ScrLen >= #Aux.DrillDepthMax)) 成立时，将 TRUE 传送到 "DB1148_PromptBeeper".Public.DrillDepthErr
   IF (((#DownDrillStep.S20 AND NOT (#DownDrillStep.S22)) AND TRUE) AND ("DB1900_Communication_PC".Send.ScrLen >= #Aux.DrillDepthMax)) THEN
       "DB1148_PromptBeeper".Public.DrillDepthErr := TRUE;
   END_IF;
   // 含义：条件 (((#DownDrillStep.S20 AND NOT (#DownDrillStep.S22)) AND "DB720_KuKa_MainCtrl".StatusIn.do_ReqStopDril) AND ("DB1900_Communication_PC".Send.ScrLen > #Aux.DrillDepthMin)) 成立时，将 0 传送到 "DB1042_Timer".DTimeOutTimes
   IF (((#DownDrillStep.S20 AND NOT (#DownDrillStep.S22)) AND "DB720_KuKa_MainCtrl".StatusIn.do_ReqStopDril) AND ("DB1900_Communication_PC".Send.ScrLen > #Aux.DrillDepthMin)) THEN
       "DB1042_Timer".DTimeOutTimes := 0;
   END_IF;
   // 含义：条件 (((((((#DownDrillStep.S20 AND NOT (#DownDrillStep.S22)) AND "DB720_KuKa_MainCtrl".StatusIn.do_DownDril_Pos) AND NOT (#DownDrillStep.StopDrill_Ack)) AND ("DB1900_Communication_PC".Recv.Current_2 > "DB1900_Communication_PC".Para.CurrentMinLimit))) AND ("DB1900_Communication_PC".Recv.Current_2 < "DB1900_Communication_PC".Para.CurrentMaxLimit))) AND "DB1042_Timer".DCurrentLastTime.Q 成立时，将 0 传送到 "DB1042_Timer".DCLowTimeOutTimes
   IF (((((((#DownDrillStep.S20 AND NOT (#DownDrillStep.S22)) AND "DB720_KuKa_MainCtrl".StatusIn.do_DownDril_Pos) AND NOT (#DownDrillStep.StopDrill_Ack)) AND ("DB1900_Communication_PC".Recv.Current_2 > "DB1900_Communication_PC".Para.CurrentMinLimit))) AND ("DB1900_Communication_PC".Recv.Current_2 < "DB1900_Communication_PC".Para.CurrentMaxLimit))) AND "DB1042_Timer".DCurrentLastTime.Q THEN
       "DB1042_Timer".DCLowTimeOutTimes := 0;
   END_IF;
   // 含义：调用计数器实例 "DB1042_Timer".DCurrentLastTime.TON（上升沿计数，当前值写入 CV）
   "DB1042_Timer".DCurrentLastTime.TON(IN := ((((((#DownDrillStep.S20 AND NOT (#DownDrillStep.S22)) AND "DB720_KuKa_MainCtrl".StatusIn.do_DownDril_Pos) AND NOT (#DownDrillStep.StopDrill_Ack)) AND ("DB1900_Communication_PC".Recv.Current_2 > "DB1900_Communication_PC".Para.CurrentMinLimit))) AND ("DB1900_Communication_PC".Recv.Current_2 < "DB1900_Communication_PC".Para.CurrentMaxLimit)),
                                       PT := T#500ms);
   // 含义：条件 ((((#DownDrillStep.S20 AND NOT (#DownDrillStep.S22)) AND "DB720_KuKa_MainCtrl".StatusIn.do_DownDril_Pos) AND #DownDrillStep.StopDrill_Ack) AND ("DB1900_Communication_PC".Send.ScrLen > #Aux.DrillDepthMin)) 成立时，将 0 传送到 "DB1042_Timer".DTimeOutTimes
   IF ((((#DownDrillStep.S20 AND NOT (#DownDrillStep.S22)) AND "DB720_KuKa_MainCtrl".StatusIn.do_DownDril_Pos) AND #DownDrillStep.StopDrill_Ack) AND ("DB1900_Communication_PC".Send.ScrLen > #Aux.DrillDepthMin)) THEN
       "DB1042_Timer".DTimeOutTimes := 0;
   END_IF;
   // 含义：条件 (#DownDrillStep.S20 AND NOT (#DownDrillStep.S22)) AND "DB1042_Timer".FixtureStuckTimeOut.Q 成立时，将 TRUE 传送到 #DownDrillStep.ErrEnd
   IF (#DownDrillStep.S20 AND NOT (#DownDrillStep.S22)) AND "DB1042_Timer".FixtureStuckTimeOut.Q THEN
       #DownDrillStep.ErrEnd := TRUE;
   END_IF;
   // 含义：条件 (#DownDrillStep.S20 AND NOT (#DownDrillStep.S22)) AND "DB1042_Timer".FixtureStuckTimeOut.Q 成立时，将 TRUE 传送到 "DB1148_PromptBeeper".Public.BitStuckErr_Fixture
   IF (#DownDrillStep.S20 AND NOT (#DownDrillStep.S22)) AND "DB1042_Timer".FixtureStuckTimeOut.Q THEN
       "DB1148_PromptBeeper".Public.BitStuckErr_Fixture := TRUE;
   END_IF;
   // 含义：条件 (#DownDrillStep.S20 AND NOT (#DownDrillStep.S22)) AND "DB1042_Timer".DrillingHighCurrentOut.Q 成立时，将 TRUE 传送到 #DownDrillStep.ErrEnd
   IF (#DownDrillStep.S20 AND NOT (#DownDrillStep.S22)) AND "DB1042_Timer".DrillingHighCurrentOut.Q THEN
       #DownDrillStep.ErrEnd := TRUE;
   END_IF;
   // 含义：条件 (#DownDrillStep.S20 AND NOT (#DownDrillStep.S22)) AND "DB1042_Timer".DrillingHighCurrentOut.Q 成立时，将 TRUE 传送到 "DB1148_PromptBeeper".Public.BitStuckErr_HighCurrent
   IF (#DownDrillStep.S20 AND NOT (#DownDrillStep.S22)) AND "DB1042_Timer".DrillingHighCurrentOut.Q THEN
       "DB1148_PromptBeeper".Public.BitStuckErr_HighCurrent := TRUE;
   END_IF;

   // ---------- 网络 20 ----------
   // 标题：TaskDone
   // 含义：条件 ((#DownDrillStep.S22 OR #DownDrillStep.ErrEnd OR #DownDrillStep.ByPass) AND NOT (#DownDrillStep.S25)) AND NOT (#DownDrillStep.ErrEnd) 成立时，将 TRUE 传送到 #DownDrillStep.TaskIO
   IF ((#DownDrillStep.S22 OR #DownDrillStep.ErrEnd OR #DownDrillStep.ByPass) AND NOT (#DownDrillStep.S25)) AND NOT (#DownDrillStep.ErrEnd) THEN
       #DownDrillStep.TaskIO := TRUE;
   END_IF;
   // 含义：条件 ((#DownDrillStep.S22 OR #DownDrillStep.ErrEnd OR #DownDrillStep.ByPass) AND NOT (#DownDrillStep.S25)) AND #DownDrillStep.ErrEnd 成立时，将 TRUE 传送到 #DownDrillStep.TaskNIO
   IF ((#DownDrillStep.S22 OR #DownDrillStep.ErrEnd OR #DownDrillStep.ByPass) AND NOT (#DownDrillStep.S25)) AND #DownDrillStep.ErrEnd THEN
       #DownDrillStep.TaskNIO := TRUE;
   END_IF;
   // 含义：条件 (#DownDrillStep.S22 OR #DownDrillStep.ErrEnd OR #DownDrillStep.ByPass) AND NOT (#DownDrillStep.S25) 成立时，将 FALSE 传送到 "DB1042_Timer".FirstStart
   IF (#DownDrillStep.S22 OR #DownDrillStep.ErrEnd OR #DownDrillStep.ByPass) AND NOT (#DownDrillStep.S25) THEN
       "DB1042_Timer".FirstStart := FALSE;
   END_IF;
   // 含义：将 #DownDrillStep.S22 OR #DownDrillStep.ErrEnd OR #DownDrillStep.ByPass 赋给 #DownDrillStep.S25
   #DownDrillStep.S25 := #DownDrillStep.S22 OR #DownDrillStep.ErrEnd OR #DownDrillStep.ByPass;

   // ---------- 网络 21 ----------
   // 标题：结束
   // 含义：将 #DownDrillStep.S25 AND NOT (#DownDrillStep.StartCmd) 赋给 #DownDrillStep.StepEnd
   #DownDrillStep.StepEnd := #DownDrillStep.S25 AND NOT (#DownDrillStep.StartCmd);
   // 含义：条件 #DownDrillStep.S25 AND #DownDrillStep.ErrEnd 成立时，将 TRUE 传送到 "DB1080_Component".Robot.Cmd.Auto.Stop
   IF #DownDrillStep.S25 AND #DownDrillStep.ErrEnd THEN
       "DB1080_Component".Robot.Cmd.Auto.Stop := TRUE;
   END_IF;
   // 含义：将 (#DownDrillStep.S25 AND "DB1080_Component".Robot.Status.TaskDone) OR (#DownDrillStep.S25 AND #DownDrillStep.TaskDone) 赋给 #DownDrillStep.TaskDone
   #DownDrillStep.TaskDone := (#DownDrillStep.S25 AND "DB1080_Component".Robot.Status.TaskDone) OR (#DownDrillStep.S25 AND #DownDrillStep.TaskDone);

   // ---------- 网络 22 ----------
   // 标题：Alarm When Drilling and  Robot Move from DownAppPos to DownInPos
   // 含义：将 FALSE 赋给 #DownDrillStep.StartCmd
   #DownDrillStep.StartCmd := FALSE;
   // 含义：条件 "DB1900_Communication_PC".Para.ProduceMode3 AND NOT ("DB720_KuKa_MainCtrl".StatusIn.do_DrilEnd_Pos) 成立时，将 FALSE 传送到 "DB1060_AutoStep".DownDrillAutoStep.DownDrillStep.ChiselEndPos
   IF "DB1900_Communication_PC".Para.ProduceMode3 AND NOT ("DB720_KuKa_MainCtrl".StatusIn.do_DrilEnd_Pos) THEN
       "DB1060_AutoStep".DownDrillAutoStep.DownDrillStep.ChiselEndPos := FALSE;
   END_IF;
END_FUNCTION_BLOCK

FUNCTION_BLOCK "FB1064_DiamondAutostep"   // FB1064, SCL
{ S7_Optimized_Access := 'TRUE' }
// ============================================================
//  Block: FB1064_DiamondAutostep
//  ============================================================
//  编号：FB1064
//  原始语言：LAD（规则翻译为 SCL）
//  含义：Water Value Control
   VAR
      Aux : Struct   // 静态变量
         OffsetX : Real;   // 静态变量
         OffsetXMid : DInt;   // 静态变量
         VibCylinderTimer : IEC_TIMER;   // 静态变量
         DiamondDetcOKTimer : IEC_TIMER;   // 静态变量
         DiamondDetcNOKTimer : IEC_TIMER;   // 静态变量
      END_STRUCT;
      EdgeDetc : Struct   // 静态变量
         Pulse : Array[0..15] of Bool;   // 静态变量
      END_STRUCT;
      DiamondStep : Struct   // 自动流程步
         Busy : Bool;   // 静态变量
         StartCmd : Bool;   // 静态变量
         OKToStart : Bool;   // 静态变量
         TaskDone : Bool;   // 静态变量
         StepStart : Bool;   // 静态变量
         StepEnd : Bool;   // 静态变量
         ErrEnd : Bool;   // 静态变量
         ByPass : Bool;   // 静态变量
         TaskIO : Bool;   // 静态变量
         TaskNIO : Bool;   // 静态变量
         S1 : Bool;   // 静态变量
         S2 : Bool;   // 静态变量
         S3 : Bool;   // 静态变量
         S4 : Bool;   // 静态变量
         S5 : Bool;   // 静态变量
         S6 : Bool;   // 静态变量
         S7 : Bool;   // 静态变量
         S8 : Bool;   // 静态变量
         S9 : Bool;   // 静态变量
         S10 : Bool;   // 静态变量
         S11 : Bool;   // 静态变量
         S12 : Bool;   // 静态变量
         S13 : Bool;   // 静态变量
         S14 : Bool;   // 静态变量
         S15 : Bool;   // 静态变量
         S16 : Bool;   // 静态变量
      END_STRUCT;
      PT : Time;   // 静态变量
      ET : Time;   // 静态变量
      IN : Bool;   // 静态变量
      Q : Bool;   // 静态变量
   END_VAR
BEGIN

   // ---------- 网络 1 ----------
   // 标题：Water Valve
   // 注释：Water Value Control
   // 含义：将 (((((("DB720_KuKa_MainCtrl".CmdOut.gi_ToolTypeNo = 13) AND "AutoMode_M") AND ("DB1900_Communication_PC".Send.ScrLen >= 6.0))) AND "DB1060_AutoStep".HorDrillAutoStep.HorDrillStep.StepStart) AND NOT ("DB1060_AutoStep".HorDrillAutoStep.HorDrillStep.StopDrill_Ack)) OR (((((("DB720_KuKa_MainCtrl".CmdOut.gi_ToolTypeNo = 13) AND "AutoMode_M") AND ("DB1900_Communication_PC".Send.ScrLen >= 6.0))) AND "DB1060_AutoStep".DownDrillAutoStep.DownDrillStep.StepStart) AND NOT ("DB1060_AutoStep".DownDrillAutoStep.DownDrillStep.StopDrill_Ack)) OR ((((("DB720_KuKa_MainCtrl".CmdOut.gi_ToolTypeNo = 13) AND "ManMode_M") AND ("DB1900_Communication_PC".Recv.Current_2 > 2.0))) AND "DB720_KuKa_MainCtrl".StatusIn.do_HorDril_Pos) OR ((((("DB720_KuKa_MainCtrl".CmdOut.gi_ToolTypeNo = 13) AND "ManMode_M") AND ("DB1900_Communication_PC".Recv.Current_2 > 2.0))) AND "DB720_KuKa_MainCtrl".StatusIn.do_DownDril_Pos) 赋给 "QWaterValve"
   "QWaterValve" := (((((("DB720_KuKa_MainCtrl".CmdOut.gi_ToolTypeNo = 13) AND "AutoMode_M") AND ("DB1900_Communication_PC".Send.ScrLen >= 6.0))) AND "DB1060_AutoStep".HorDrillAutoStep.HorDrillStep.StepStart) AND NOT ("DB1060_AutoStep".HorDrillAutoStep.HorDrillStep.StopDrill_Ack)) OR (((((("DB720_KuKa_MainCtrl".CmdOut.gi_ToolTypeNo = 13) AND "AutoMode_M") AND ("DB1900_Communication_PC".Send.ScrLen >= 6.0))) AND "DB1060_AutoStep".DownDrillAutoStep.DownDrillStep.StepStart) AND NOT ("DB1060_AutoStep".DownDrillAutoStep.DownDrillStep.StopDrill_Ack)) OR ((((("DB720_KuKa_MainCtrl".CmdOut.gi_ToolTypeNo = 13) AND "ManMode_M") AND ("DB1900_Communication_PC".Recv.Current_2 > 2.0))) AND "DB720_KuKa_MainCtrl".StatusIn.do_HorDril_Pos) OR ((((("DB720_KuKa_MainCtrl".CmdOut.gi_ToolTypeNo = 13) AND "ManMode_M") AND ("DB1900_Communication_PC".Recv.Current_2 > 2.0))) AND "DB720_KuKa_MainCtrl".StatusIn.do_DownDril_Pos);
   // 含义：条件 (((((("DB720_KuKa_MainCtrl".CmdOut.gi_ToolTypeNo = 13) AND "AutoMode_M") AND "DB1060_AutoStep".HorDrillAutoStep.Aux.StartDrill) AND NOT ("DB1060_AutoStep".HorDrillAutoStep.HorDrillStep.StopDrill_Ack)) OR (((("DB720_KuKa_MainCtrl".CmdOut.gi_ToolTypeNo = 13) AND "AutoMode_M") AND "DB1060_AutoStep".DownDrillAutoStep.Aux.StartDrill) AND NOT ("DB1060_AutoStep".DownDrillAutoStep.DownDrillStep.StopDrill_Ack))) AND ("DB1900_Communication_PC".Send.ScrLen < 10.0)) 成立时，将 2 传送到 "DB1080_Component".Robot.CTRL_IN.RobotSpeed
   IF (((((("DB720_KuKa_MainCtrl".CmdOut.gi_ToolTypeNo = 13) AND "AutoMode_M") AND "DB1060_AutoStep".HorDrillAutoStep.Aux.StartDrill) AND NOT ("DB1060_AutoStep".HorDrillAutoStep.HorDrillStep.StopDrill_Ack)) OR (((("DB720_KuKa_MainCtrl".CmdOut.gi_ToolTypeNo = 13) AND "AutoMode_M") AND "DB1060_AutoStep".DownDrillAutoStep.Aux.StartDrill) AND NOT ("DB1060_AutoStep".DownDrillAutoStep.DownDrillStep.StopDrill_Ack))) AND ("DB1900_Communication_PC".Send.ScrLen < 10.0)) THEN
       "DB1080_Component".Robot.CTRL_IN.RobotSpeed := 2;
   END_IF;
   // 含义：条件 ((((((("DB720_KuKa_MainCtrl".CmdOut.gi_ToolTypeNo = 13) AND "AutoMode_M") AND "DB1060_AutoStep".HorDrillAutoStep.Aux.StartDrill) AND NOT ("DB1060_AutoStep".HorDrillAutoStep.HorDrillStep.StopDrill_Ack)) OR (((("DB720_KuKa_MainCtrl".CmdOut.gi_ToolTypeNo = 13) AND "AutoMode_M") AND "DB1060_AutoStep".DownDrillAutoStep.Aux.StartDrill) AND NOT ("DB1060_AutoStep".DownDrillAutoStep.DownDrillStep.StopDrill_Ack))) AND ("DB1900_Communication_PC".Send.ScrLen >= 10.0))) AND TRUE 成立时，将 FALSE 传送到 "QCamCoverExt"
   IF ((((((("DB720_KuKa_MainCtrl".CmdOut.gi_ToolTypeNo = 13) AND "AutoMode_M") AND "DB1060_AutoStep".HorDrillAutoStep.Aux.StartDrill) AND NOT ("DB1060_AutoStep".HorDrillAutoStep.HorDrillStep.StopDrill_Ack)) OR (((("DB720_KuKa_MainCtrl".CmdOut.gi_ToolTypeNo = 13) AND "AutoMode_M") AND "DB1060_AutoStep".DownDrillAutoStep.Aux.StartDrill) AND NOT ("DB1060_AutoStep".DownDrillAutoStep.DownDrillStep.StopDrill_Ack))) AND ("DB1900_Communication_PC".Send.ScrLen >= 10.0))) AND TRUE THEN
       "QCamCoverExt" := FALSE;
   END_IF;
   // 含义：条件 ((((((("DB720_KuKa_MainCtrl".CmdOut.gi_ToolTypeNo = 13) AND "AutoMode_M") AND "DB1060_AutoStep".HorDrillAutoStep.Aux.StartDrill) AND NOT ("DB1060_AutoStep".HorDrillAutoStep.HorDrillStep.StopDrill_Ack)) OR (((("DB720_KuKa_MainCtrl".CmdOut.gi_ToolTypeNo = 13) AND "AutoMode_M") AND "DB1060_AutoStep".DownDrillAutoStep.Aux.StartDrill) AND NOT ("DB1060_AutoStep".DownDrillAutoStep.DownDrillStep.StopDrill_Ack))) AND ("DB1900_Communication_PC".Send.ScrLen >= 10.0))) AND TRUE 成立时，将 FALSE 传送到 "QCamCoverRet"
   IF ((((((("DB720_KuKa_MainCtrl".CmdOut.gi_ToolTypeNo = 13) AND "AutoMode_M") AND "DB1060_AutoStep".HorDrillAutoStep.Aux.StartDrill) AND NOT ("DB1060_AutoStep".HorDrillAutoStep.HorDrillStep.StopDrill_Ack)) OR (((("DB720_KuKa_MainCtrl".CmdOut.gi_ToolTypeNo = 13) AND "AutoMode_M") AND "DB1060_AutoStep".DownDrillAutoStep.Aux.StartDrill) AND NOT ("DB1060_AutoStep".DownDrillAutoStep.DownDrillStep.StopDrill_Ack))) AND ("DB1900_Communication_PC".Send.ScrLen >= 10.0))) AND TRUE THEN
       "QCamCoverRet" := FALSE;
   END_IF;
   // InRange resolved: 10.0 <= ScrLen <= 20.0
   IF ("DB1900_Communication_PC".Para.RobotSpeed >= 6.0 AND "DB1900_Communication_PC".Para.RobotSpeed <= 9.0) THEN
       "DB1080_Component".Robot.CTRL_IN.RobotSpeed := 4;
   END_IF;
   IF ("DB1900_Communication_PC".Para.RobotSpeed >= 10.0 AND "DB1900_Communication_PC".Para.RobotSpeed <= 14.0) THEN
       "DB1080_Component".Robot.CTRL_IN.RobotSpeed := 6;
   END_IF;
   IF ("DB1900_Communication_PC".Para.RobotSpeed >= 15.0 AND "DB1900_Communication_PC".Para.RobotSpeed <= 20.0) THEN
       "DB1080_Component".Robot.CTRL_IN.RobotSpeed := 8;
   END_IF;
   // 含义：条件 ("DB1900_Communication_PC".Para.RobotSpeed > 20.0) 成立时，将 10 传送到 "DB1080_Component".Robot.CTRL_IN.RobotSpeed
   IF ("DB1900_Communication_PC".Para.RobotSpeed > 20.0) THEN
       "DB1080_Component".Robot.CTRL_IN.RobotSpeed := 10;
   END_IF;

   // ---------- 网络 2 ----------
   // 标题：本工位必须要做(可能条件暂时不满足)
   // 含义：将 (("DB720_KuKa_MainCtrl".Ctrl_Out.RobotAction = 0) AND "DB720_KuKa_MainCtrl".Aux.ToolAtPos) AND NOT ("DB1148_PromptBeeper".Public.RobotNotReady) 赋给 #DiamondStep.OKToStart
   #DiamondStep.OKToStart := (("DB720_KuKa_MainCtrl".Ctrl_Out.RobotAction = 0) AND "DB720_KuKa_MainCtrl".Aux.ToolAtPos) AND NOT ("DB1148_PromptBeeper".Public.RobotNotReady);

   // ---------- 网络 3 ----------
   // 标题：*********************************岩芯去除Start****************************************
   // 含义：将 ((((((((#DiamondStep.StartCmd AND #DiamondStep.OKToStart) OR #DiamondStep.StepStart) AND "AllMode_M") AND NOT ("DB1040_HomePos".Status.Running)) AND NOT ("DB1900_Communication_PC".Recv.EmmMode)) AND ("DB720_KuKa_MainCtrl".CmdOut.gi_ToolTypeNo <> 2))) AND NOT (#DiamondStep.StepEnd)) AND NOT (#DiamondStep.ErrEnd) 赋给 #DiamondStep.StepStart
   #DiamondStep.StepStart := ((((((((#DiamondStep.StartCmd AND #DiamondStep.OKToStart) OR #DiamondStep.StepStart) AND "AllMode_M") AND NOT ("DB1040_HomePos".Status.Running)) AND NOT ("DB1900_Communication_PC".Recv.EmmMode)) AND ("DB720_KuKa_MainCtrl".CmdOut.gi_ToolTypeNo <> 2))) AND NOT (#DiamondStep.StepEnd)) AND NOT (#DiamondStep.ErrEnd);
   // 含义：条件 NOT (((((((((#DiamondStep.StartCmd AND #DiamondStep.OKToStart) OR #DiamondStep.StepStart) AND "AllMode_M") AND NOT ("DB1040_HomePos".Status.Running)) AND NOT ("DB1900_Communication_PC".Recv.EmmMode)) AND ("DB720_KuKa_MainCtrl".CmdOut.gi_ToolTypeNo <> 2))) AND NOT (#DiamondStep.StepEnd)) AND NOT (#DiamondStep.ErrEnd)) 成立时，将 FALSE 传送到 #DiamondStep.ErrEnd
   IF NOT (((((((((#DiamondStep.StartCmd AND #DiamondStep.OKToStart) OR #DiamondStep.StepStart) AND "AllMode_M") AND NOT ("DB1040_HomePos".Status.Running)) AND NOT ("DB1900_Communication_PC".Recv.EmmMode)) AND ("DB720_KuKa_MainCtrl".CmdOut.gi_ToolTypeNo <> 2))) AND NOT (#DiamondStep.StepEnd)) AND NOT (#DiamondStep.ErrEnd)) THEN
       #DiamondStep.ErrEnd := FALSE;
   END_IF;
   // 含义：条件 NOT (((((((((#DiamondStep.StartCmd AND #DiamondStep.OKToStart) OR #DiamondStep.StepStart) AND "AllMode_M") AND NOT ("DB1040_HomePos".Status.Running)) AND NOT ("DB1900_Communication_PC".Recv.EmmMode)) AND ("DB720_KuKa_MainCtrl".CmdOut.gi_ToolTypeNo <> 2))) AND NOT (#DiamondStep.StepEnd)) AND NOT (#DiamondStep.ErrEnd)) 成立时，将 FALSE 传送到 "DiamondVibCylinder"
   IF NOT (((((((((#DiamondStep.StartCmd AND #DiamondStep.OKToStart) OR #DiamondStep.StepStart) AND "AllMode_M") AND NOT ("DB1040_HomePos".Status.Running)) AND NOT ("DB1900_Communication_PC".Recv.EmmMode)) AND ("DB720_KuKa_MainCtrl".CmdOut.gi_ToolTypeNo <> 2))) AND NOT (#DiamondStep.StepEnd)) AND NOT (#DiamondStep.ErrEnd)) THEN
       "DiamondVibCylinder" := FALSE;
   END_IF;
   // 含义：条件 NOT (((((((((#DiamondStep.StartCmd AND #DiamondStep.OKToStart) OR #DiamondStep.StepStart) AND "AllMode_M") AND NOT ("DB1040_HomePos".Status.Running)) AND NOT ("DB1900_Communication_PC".Recv.EmmMode)) AND ("DB720_KuKa_MainCtrl".CmdOut.gi_ToolTypeNo <> 2))) AND NOT (#DiamondStep.StepEnd)) AND NOT (#DiamondStep.ErrEnd)) 成立时，将 FALSE 传送到 "DB720_KuKa_MainCtrl".CmdOut.di_DiamondVib_Ack
   IF NOT (((((((((#DiamondStep.StartCmd AND #DiamondStep.OKToStart) OR #DiamondStep.StepStart) AND "AllMode_M") AND NOT ("DB1040_HomePos".Status.Running)) AND NOT ("DB1900_Communication_PC".Recv.EmmMode)) AND ("DB720_KuKa_MainCtrl".CmdOut.gi_ToolTypeNo <> 2))) AND NOT (#DiamondStep.StepEnd)) AND NOT (#DiamondStep.ErrEnd)) THEN
       "DB720_KuKa_MainCtrl".CmdOut.di_DiamondVib_Ack := FALSE;
   END_IF;

   // ---------- 网络 4 ----------
   // 标题：初始化
   // 注释：Added DB2700.VisualChiselingStart  by WXY, 20220615.
   // 含义：条件 (#DiamondStep.StepStart AND NOT (#DiamondStep.ErrEnd)) AND NOT (#DiamondStep.S1) 成立时，将 FALSE 传送到 #DiamondStep.TaskIO
   IF (#DiamondStep.StepStart AND NOT (#DiamondStep.ErrEnd)) AND NOT (#DiamondStep.S1) THEN
       #DiamondStep.TaskIO := FALSE;
   END_IF;
   // 含义：条件 (#DiamondStep.StepStart AND NOT (#DiamondStep.ErrEnd)) AND NOT (#DiamondStep.S1) 成立时，将 FALSE 传送到 #DiamondStep.TaskNIO
   IF (#DiamondStep.StepStart AND NOT (#DiamondStep.ErrEnd)) AND NOT (#DiamondStep.S1) THEN
       #DiamondStep.TaskNIO := FALSE;
   END_IF;
   // 含义：将 #DiamondStep.StepStart AND NOT (#DiamondStep.ErrEnd) 赋给 #DiamondStep.S1
   #DiamondStep.S1 := #DiamondStep.StepStart AND NOT (#DiamondStep.ErrEnd);
   // 含义：将 ((((#DiamondStep.StepStart AND NOT (#DiamondStep.ErrEnd)) AND ("DB720_KuKa_MainCtrl".CmdOut.gi_ToolTypeNo = 18))) AND ("DB1900_Communication_PC".Para.DrillDepth < 100.0)) 赋给 "DB720_KuKa_MainCtrl".CmdOut.di_NotDectceDiamond
   "DB720_KuKa_MainCtrl".CmdOut.di_NotDectceDiamond := ((((#DiamondStep.StepStart AND NOT (#DiamondStep.ErrEnd)) AND ("DB720_KuKa_MainCtrl".CmdOut.gi_ToolTypeNo = 18))) AND ("DB1900_Communication_PC".Para.DrillDepth < 100.0));

   // ---------- 网络 5 ----------
   // 标题：初始化气缸
   // 含义：条件 #DiamondStep.S1 AND NOT (#DiamondStep.S3) 成立时，将 TRUE 传送到 "DB1081_ValveCall".ST01.Z01.ExtAuto
   IF #DiamondStep.S1 AND NOT (#DiamondStep.S3) THEN
       "DB1081_ValveCall".ST01.Z01.ExtAuto := TRUE;
   END_IF;
   // 含义：条件 #DiamondStep.S1 AND NOT (#DiamondStep.S3) 成立时，将 TRUE 传送到 "DB1081_ValveCall".ST01.Z02.VentValveAuto
   IF #DiamondStep.S1 AND NOT (#DiamondStep.S3) THEN
       "DB1081_ValveCall".ST01.Z02.VentValveAuto := TRUE;
   END_IF;
   // 含义：条件 (#DiamondStep.S1 AND NOT (#DiamondStep.S3)) AND TRUE 成立时，将 FALSE 传送到 "QCamCoverExt"
   IF (#DiamondStep.S1 AND NOT (#DiamondStep.S3)) AND TRUE THEN
       "QCamCoverExt" := FALSE;
   END_IF;
   // 含义：条件 (#DiamondStep.S1 AND NOT (#DiamondStep.S3)) AND TRUE 成立时，将 TRUE 传送到 "QCamCoverRet"
   IF (#DiamondStep.S1 AND NOT (#DiamondStep.S3)) AND TRUE THEN
       "QCamCoverRet" := TRUE;
   END_IF;
   // 含义：条件 #DiamondStep.S1 AND NOT (#DiamondStep.S3) 成立时，将 TRUE 传送到 "DB1081_ValveCall".ST01.Z05.RetAuto
   IF #DiamondStep.S1 AND NOT (#DiamondStep.S3) THEN
       "DB1081_ValveCall".ST01.Z05.RetAuto := TRUE;
   END_IF;
   // 含义：条件 #DiamondStep.S1 AND NOT (#DiamondStep.S3) 成立时，将 0.45 传送到 "DB1080_Component".Aux.Pressure
   IF #DiamondStep.S1 AND NOT (#DiamondStep.S3) THEN
       "DB1080_Component".Aux.Pressure := 0.45;
   END_IF;
   // 含义：将 (#DiamondStep.S1 AND "DB1081_ValveCall".ST01.Z05.IRetPos) OR (#DiamondStep.S1 AND #DiamondStep.S3) 赋给 #DiamondStep.S3
   #DiamondStep.S3 := (#DiamondStep.S1 AND "DB1081_ValveCall".ST01.Z05.IRetPos) OR (#DiamondStep.S1 AND #DiamondStep.S3);

   // ---------- 网络 6 ----------
   // 标题：偏移计算
   // 注释：示教基准为32mm钻头
   // 32mm: Hor; Heiggt:  45mm;
   // 52mm:Down; Height: 65mm;
   // 82mm Hor; Height: 90mm;
   // 102mm Hor; Height: 80mm;
   // 132mm Hor; Height: 120mm;
   // 含义：条件 ((((#DiamondStep.S3 AND NOT (#DiamondStep.S5)) AND ("DB720_KuKa_MainCtrl".CmdOut.gi_ToolTypeNo = 13))) AND ("DB1900_Communication_PC".Para.DrillWidth = 45.0)) 成立时，将 (32.0-32.0)/ 2.0 传送到 #Aux.OffsetX
   IF ((((#DiamondStep.S3 AND NOT (#DiamondStep.S5)) AND ("DB720_KuKa_MainCtrl".CmdOut.gi_ToolTypeNo = 13))) AND ("DB1900_Communication_PC".Para.DrillWidth = 45.0)) THEN
       #Aux.OffsetX := (32.0 - 32.0) / 2.0;
   END_IF;
   // 含义：条件 ((((#DiamondStep.S3 AND NOT (#DiamondStep.S5)) AND ("DB720_KuKa_MainCtrl".CmdOut.gi_ToolTypeNo = 13))) AND ("DB1900_Communication_PC".Para.DrillWidth = 65.0)) 成立时，将 (52.0-32.0)/ 2.0 传送到 #Aux.OffsetX
   IF ((((#DiamondStep.S3 AND NOT (#DiamondStep.S5)) AND ("DB720_KuKa_MainCtrl".CmdOut.gi_ToolTypeNo = 13))) AND ("DB1900_Communication_PC".Para.DrillWidth = 65.0)) THEN
       #Aux.OffsetX := (52.0 - 32.0) / 2.0;
   END_IF;
   // 含义：条件 ((((#DiamondStep.S3 AND NOT (#DiamondStep.S5)) AND ("DB720_KuKa_MainCtrl".CmdOut.gi_ToolTypeNo = 13))) AND ("DB1900_Communication_PC".Para.DrillWidth = 85.0)) 成立时，将 (82.0-32.0)/ 2.0 传送到 #Aux.OffsetX
   IF ((((#DiamondStep.S3 AND NOT (#DiamondStep.S5)) AND ("DB720_KuKa_MainCtrl".CmdOut.gi_ToolTypeNo = 13))) AND ("DB1900_Communication_PC".Para.DrillWidth = 85.0)) THEN
       #Aux.OffsetX := (82.0 - 32.0) / 2.0;
   END_IF;
   // 含义：条件 ((((#DiamondStep.S3 AND NOT (#DiamondStep.S5)) AND ("DB720_KuKa_MainCtrl".CmdOut.gi_ToolTypeNo = 13))) AND ("DB1900_Communication_PC".Para.DrillWidth = 80.0)) 成立时，将 (102.0-32.0)/ 2.0 传送到 #Aux.OffsetX
   IF ((((#DiamondStep.S3 AND NOT (#DiamondStep.S5)) AND ("DB720_KuKa_MainCtrl".CmdOut.gi_ToolTypeNo = 13))) AND ("DB1900_Communication_PC".Para.DrillWidth = 80.0)) THEN
       #Aux.OffsetX := (102.0 - 32.0) / 2.0;
   END_IF;
   // 含义：条件 ((((#DiamondStep.S3 AND NOT (#DiamondStep.S5)) AND ("DB720_KuKa_MainCtrl".CmdOut.gi_ToolTypeNo = 13))) AND ("DB1900_Communication_PC".Para.DrillWidth = 120.0)) 成立时，将 (132.0-32.0)/ 2.0 传送到 #Aux.OffsetX
   IF ((((#DiamondStep.S3 AND NOT (#DiamondStep.S5)) AND ("DB720_KuKa_MainCtrl".CmdOut.gi_ToolTypeNo = 13))) AND ("DB1900_Communication_PC".Para.DrillWidth = 120.0)) THEN
       #Aux.OffsetX := (132.0 - 32.0) / 2.0;
   END_IF;
   // 含义：条件 ((((#DiamondStep.S3 AND NOT (#DiamondStep.S5)) AND ("DB720_KuKa_MainCtrl".CmdOut.gi_ToolTypeNo = 18))) AND ("DB1900_Communication_PC".Para.DrillWidth = 90.0)) 成立时，将 5.0 传送到 #Aux.OffsetX
   IF ((((#DiamondStep.S3 AND NOT (#DiamondStep.S5)) AND ("DB720_KuKa_MainCtrl".CmdOut.gi_ToolTypeNo = 18))) AND ("DB1900_Communication_PC".Para.DrillWidth = 90.0)) THEN
       #Aux.OffsetX := 5.0;
   END_IF;
   // 含义：条件 ((((#DiamondStep.S3 AND NOT (#DiamondStep.S5)) AND ("DB720_KuKa_MainCtrl".CmdOut.gi_ToolTypeNo = 18))) AND ("DB1900_Communication_PC".Para.DrillWidth = 80.0)) 成立时，将 0.0 传送到 #Aux.OffsetX
   IF ((((#DiamondStep.S3 AND NOT (#DiamondStep.S5)) AND ("DB720_KuKa_MainCtrl".CmdOut.gi_ToolTypeNo = 18))) AND ("DB1900_Communication_PC".Para.DrillWidth = 80.0)) THEN
       #Aux.OffsetX := 0.0;
   END_IF;
   // 含义：将 #Aux.OffsetX; (* Convert → DInt *) END_IF 赋给 IF #DiamondStep.S3 AND NOT (#DiamondStep.S5) THEN #Aux.OffsetXMid
   IF #DiamondStep.S3 AND NOT (#DiamondStep.S5) THEN
       #Aux.OffsetXMid := #Aux.OffsetX; (* Convert → DInt *)
   END_IF;
   // 含义：将 SWAP(#Aux.OffsetXMid) 赋给 "DB720_KuKa_MainCtrl".CmdOut.gi_OffSetX
   "DB720_KuKa_MainCtrl".CmdOut.gi_OffSetX := SWAP(#Aux.OffsetXMid);
   // 含义：当 #DiamondStep.S3 为 TRUE 时置位 #DiamondStep.S5，否则复位（触点→线圈）
   IF #DiamondStep.S3 THEN
       #DiamondStep.S5 := TRUE;
   ELSE
       #DiamondStep.S5 := FALSE;
   END_IF;

   // ---------- 网络 7 ----------
   // 含义：将 (#DiamondStep.S5 AND NOT ("DB1080_Component".Robot.Status.Busy)) OR (#DiamondStep.S5 AND #DiamondStep.S6) 赋给 #DiamondStep.S6
   #DiamondStep.S6 := (#DiamondStep.S5 AND NOT ("DB1080_Component".Robot.Status.Busy)) OR (#DiamondStep.S5 AND #DiamondStep.S6);

   // ---------- 网络 8 ----------
   // 标题：枪电源
   // 含义：条件 #DiamondStep.S6 AND NOT (#DiamondStep.S7) 成立时，将 17 传送到 "DB1080_Component".Robot.CTRL_IN.ProgNo
   IF #DiamondStep.S6 AND NOT (#DiamondStep.S7) THEN
       "DB1080_Component".Robot.CTRL_IN.ProgNo := 17;
   END_IF;
   // 含义：条件 #DiamondStep.S6 AND NOT (#DiamondStep.S7) 成立时，将 60 传送到 "DB1080_Component".Robot.CTRL_IN.RobotSpeed
   IF #DiamondStep.S6 AND NOT (#DiamondStep.S7) THEN
       "DB1080_Component".Robot.CTRL_IN.RobotSpeed := 60;
   END_IF;
   // 含义：条件 (((#DiamondStep.S6 AND ("DB720_KuKa_MainCtrl".CmdOut.gi_ToolTypeNo = 13))) AND "DB720_KuKa_MainCtrl".StatusIn.do_Diamond_Act) AND "DB720_KuKa_MainCtrl".StatusIn.do_JDiamond_MidPos 成立时，将 TRUE 传送到 "DB1081_ValveCall".ST01.Z05.ExtAuto
   IF (((#DiamondStep.S6 AND ("DB720_KuKa_MainCtrl".CmdOut.gi_ToolTypeNo = 13))) AND "DB720_KuKa_MainCtrl".StatusIn.do_Diamond_Act) AND "DB720_KuKa_MainCtrl".StatusIn.do_JDiamond_MidPos THEN
       "DB1081_ValveCall".ST01.Z05.ExtAuto := TRUE;
   END_IF;
   // 含义：条件 (((#DiamondStep.S6 AND ("DB720_KuKa_MainCtrl".CmdOut.gi_ToolTypeNo = 13))) AND "DB720_KuKa_MainCtrl".StatusIn.do_Diamond_Act) AND NOT ("DB720_KuKa_MainCtrl".StatusIn.do_JDiamond_MidPos) 成立时，将 TRUE 传送到 "DB1081_ValveCall".ST01.Z05.RetAuto
   IF (((#DiamondStep.S6 AND ("DB720_KuKa_MainCtrl".CmdOut.gi_ToolTypeNo = 13))) AND "DB720_KuKa_MainCtrl".StatusIn.do_Diamond_Act) AND NOT ("DB720_KuKa_MainCtrl".StatusIn.do_JDiamond_MidPos) THEN
       "DB1081_ValveCall".ST01.Z05.RetAuto := TRUE;
   END_IF;
   // 含义：条件 #DiamondStep.S6 成立时，将 TRUE 传送到 "DB1080_Component".Robot.Cmd.Auto.ProgStart
   IF #DiamondStep.S6 THEN
       "DB1080_Component".Robot.Cmd.Auto.ProgStart := TRUE;
   END_IF;
   // 含义：将 (#DiamondStep.S6 AND "DB720_KuKa_MainCtrl".StatusIn.do_Diamond_Act) OR (#DiamondStep.S6 AND #DiamondStep.S7) 赋给 #DiamondStep.S7
   #DiamondStep.S7 := (#DiamondStep.S6 AND "DB720_KuKa_MainCtrl".StatusIn.do_Diamond_Act) OR (#DiamondStep.S6 AND #DiamondStep.S7);

   // ---------- 网络 9 ----------
   // 标题：水钻振动气缸
   // 含义：条件 (((#DiamondStep.S7 AND NOT (#DiamondStep.S9)) AND ("DB1900_Communication_PC".Recv.Current_2 < 1.0))) AND "DB720_KuKa_MainCtrl".StatusIn.do_DiamondVib_Pos 成立时，将 TRUE 传送到 "DiamondVibCylinder"
   IF (((#DiamondStep.S7 AND NOT (#DiamondStep.S9)) AND ("DB1900_Communication_PC".Recv.Current_2 < 1.0))) AND "DB720_KuKa_MainCtrl".StatusIn.do_DiamondVib_Pos THEN
       "DiamondVibCylinder" := TRUE;
   END_IF;
   // 含义：调用计数器实例 #Aux.VibCylinderTimer.TON（上升沿计数，当前值写入 CV）
   #Aux.VibCylinderTimer.TON(IN := (((#DiamondStep.S7 AND NOT (#DiamondStep.S9)) AND ("DB1900_Communication_PC".Recv.Current_2 < 1.0))) AND "DiamondVibCylinder",
                             PT := T#3S);
   // 含义：条件 (((#DiamondStep.S7 AND NOT (#DiamondStep.S9)) AND ("DB1900_Communication_PC".Recv.Current_2 < 1.0))) AND #Aux.VibCylinderTimer.Q 成立时，将 FALSE 传送到 "DiamondVibCylinder"
   IF (((#DiamondStep.S7 AND NOT (#DiamondStep.S9)) AND ("DB1900_Communication_PC".Recv.Current_2 < 1.0))) AND #Aux.VibCylinderTimer.Q THEN
       "DiamondVibCylinder" := FALSE;
   END_IF;
   // 含义：条件 (((#DiamondStep.S7 AND NOT (#DiamondStep.S9)) AND ("DB1900_Communication_PC".Recv.Current_2 < 1.0))) AND #Aux.VibCylinderTimer.Q 成立时，将 TRUE 传送到 "DB720_KuKa_MainCtrl".CmdOut.di_DiamondVib_Ack
   IF (((#DiamondStep.S7 AND NOT (#DiamondStep.S9)) AND ("DB1900_Communication_PC".Recv.Current_2 < 1.0))) AND #Aux.VibCylinderTimer.Q THEN
       "DB720_KuKa_MainCtrl".CmdOut.di_DiamondVib_Ack := TRUE;
   END_IF;
   // 含义：将 (#DiamondStep.S7 AND #Aux.VibCylinderTimer.Q) OR (#DiamondStep.S7 AND #DiamondStep.S9) 赋给 #DiamondStep.S9
   #DiamondStep.S9 := (#DiamondStep.S7 AND #Aux.VibCylinderTimer.Q) OR (#DiamondStep.S7 AND #DiamondStep.S9);

   // ---------- 网络 10 ----------
   // 标题：岩芯检测信号
   // 含义：将 NOT ("ICoreBlockDect_LeftTool") AND NOT ("ICoreBlockDect_RightTool") 赋给 #EdgeDetc.Pulse[0]
   #EdgeDetc.Pulse[0] := NOT ("ICoreBlockDect_LeftTool") AND NOT ("ICoreBlockDect_RightTool");
   // 含义：将 NOT (NOT ("ICoreBlockDect_LeftTool") AND NOT ("ICoreBlockDect_RightTool")) 赋给 #EdgeDetc.Pulse[0]
   #EdgeDetc.Pulse[0] := NOT (NOT ("ICoreBlockDect_LeftTool") AND NOT ("ICoreBlockDect_RightTool"));
   // 含义：当 NOT ("ICoreBlockDect_LeftTool") 为 TRUE 时置位 #EdgeDetc.Pulse[0]，否则复位（触点→线圈）
   IF NOT ("ICoreBlockDect_LeftTool") THEN
       #EdgeDetc.Pulse[0] := TRUE;
   ELSE
       #EdgeDetc.Pulse[0] := FALSE;
   END_IF;
   // 含义：当 "ICoreBlockDect_LeftTool" 为 TRUE 时置位 #EdgeDetc.Pulse[0]，否则复位（触点→线圈）
   IF "ICoreBlockDect_LeftTool" THEN
       #EdgeDetc.Pulse[0] := TRUE;
   ELSE
       #EdgeDetc.Pulse[0] := FALSE;
   END_IF;

   // ---------- 网络 11 ----------
   // 标题：水钻岩芯敲击完成确认
   // 含义：调用定时器实例 #Aux.DiamondDetcOKTimer.TON
   #Aux.DiamondDetcOKTimer.TON(IN := ((((((#DiamondStep.S9 AND NOT ("DB720_KuKa_MainCtrl".CmdOut.di_NotDectceDiamond)) AND NOT (#DiamondStep.S11)) AND "DB720_KuKa_MainCtrl".StatusIn.do_DiamondDetc_Pos) AND ("DB720_KuKa_MainCtrl".CmdOut.gi_ToolTypeNo = 13))) AND #EdgeDetc.Pulse[0]) OR ((((((#DiamondStep.S9 AND NOT ("DB720_KuKa_MainCtrl".CmdOut.di_NotDectceDiamond)) AND NOT (#DiamondStep.S11)) AND "DB720_KuKa_MainCtrl".StatusIn.do_DiamondDetc_Pos) AND ("DB720_KuKa_MainCtrl".CmdOut.gi_ToolTypeNo = 18))) AND #EdgeDetc.Pulse[0]),
                               PT := T#3S);
   // 含义：条件 ((((((#DiamondStep.S9 AND NOT ("DB720_KuKa_MainCtrl".CmdOut.di_NotDectceDiamond)) AND NOT (#DiamondStep.S11)) AND "DB720_KuKa_MainCtrl".StatusIn.do_DiamondDetc_Pos) AND ("DB720_KuKa_MainCtrl".CmdOut.gi_ToolTypeNo = 13))) AND #EdgeDetc.Pulse[0]) OR ((((((#DiamondStep.S9 AND NOT ("DB720_KuKa_MainCtrl".CmdOut.di_NotDectceDiamond)) AND NOT (#DiamondStep.S11)) AND "DB720_KuKa_MainCtrl".StatusIn.do_DiamondDetc_Pos) AND ("DB720_KuKa_MainCtrl".CmdOut.gi_ToolTypeNo = 18))) AND #EdgeDetc.Pulse[0]) 成立时，将 FALSE 传送到 "DB720_KuKa_MainCtrl".CmdOut.di_DiamondVib_Ack
   IF ((((((#DiamondStep.S9 AND NOT ("DB720_KuKa_MainCtrl".CmdOut.di_NotDectceDiamond)) AND NOT (#DiamondStep.S11)) AND "DB720_KuKa_MainCtrl".StatusIn.do_DiamondDetc_Pos) AND ("DB720_KuKa_MainCtrl".CmdOut.gi_ToolTypeNo = 13))) AND #EdgeDetc.Pulse[0]) OR ((((((#DiamondStep.S9 AND NOT ("DB720_KuKa_MainCtrl".CmdOut.di_NotDectceDiamond)) AND NOT (#DiamondStep.S11)) AND "DB720_KuKa_MainCtrl".StatusIn.do_DiamondDetc_Pos) AND ("DB720_KuKa_MainCtrl".CmdOut.gi_ToolTypeNo = 18))) AND #EdgeDetc.Pulse[0]) THEN
       "DB720_KuKa_MainCtrl".CmdOut.di_DiamondVib_Ack := FALSE;
   END_IF;
   // 含义：调用定时器实例 #Aux.DiamondDetcNOKTimer.TON
   #Aux.DiamondDetcNOKTimer.TON(IN := ((((((#DiamondStep.S9 AND NOT ("DB720_KuKa_MainCtrl".CmdOut.di_NotDectceDiamond)) AND NOT (#DiamondStep.S11)) AND "DB720_KuKa_MainCtrl".StatusIn.do_DiamondDetc_Pos) AND ("DB720_KuKa_MainCtrl".CmdOut.gi_ToolTypeNo = 13))) AND #EdgeDetc.Pulse[0]) OR ((((((#DiamondStep.S9 AND NOT ("DB720_KuKa_MainCtrl".CmdOut.di_NotDectceDiamond)) AND NOT (#DiamondStep.S11)) AND "DB720_KuKa_MainCtrl".StatusIn.do_DiamondDetc_Pos) AND ("DB720_KuKa_MainCtrl".CmdOut.gi_ToolTypeNo = 18))) AND #EdgeDetc.Pulse[0]),
                                PT := T#4S);
   // 含义：条件 (((#DiamondStep.S9 AND NOT ("DB720_KuKa_MainCtrl".CmdOut.di_NotDectceDiamond)) AND NOT (#DiamondStep.S11)) AND "DB720_KuKa_MainCtrl".StatusIn.do_DiamondDetc_Pos) AND #Aux.DiamondDetcNOKTimer.Q 成立时，将 TRUE 传送到 #DiamondStep.ErrEnd
   IF (((#DiamondStep.S9 AND NOT ("DB720_KuKa_MainCtrl".CmdOut.di_NotDectceDiamond)) AND NOT (#DiamondStep.S11)) AND "DB720_KuKa_MainCtrl".StatusIn.do_DiamondDetc_Pos) AND #Aux.DiamondDetcNOKTimer.Q THEN
       #DiamondStep.ErrEnd := TRUE;
   END_IF;
   // 含义：条件 (((#DiamondStep.S9 AND NOT ("DB720_KuKa_MainCtrl".CmdOut.di_NotDectceDiamond)) AND NOT (#DiamondStep.S11)) AND "DB720_KuKa_MainCtrl".StatusIn.do_DiamondDetc_Pos) AND #Aux.DiamondDetcNOKTimer.Q 成立时，将 TRUE 传送到 "DB1080_Component".Robot.Cmd.Auto.Stop
   IF (((#DiamondStep.S9 AND NOT ("DB720_KuKa_MainCtrl".CmdOut.di_NotDectceDiamond)) AND NOT (#DiamondStep.S11)) AND "DB720_KuKa_MainCtrl".StatusIn.do_DiamondDetc_Pos) AND #Aux.DiamondDetcNOKTimer.Q THEN
       "DB1080_Component".Robot.Cmd.Auto.Stop := TRUE;
   END_IF;
   // 含义：条件 (((#DiamondStep.S9 AND NOT ("DB720_KuKa_MainCtrl".CmdOut.di_NotDectceDiamond)) AND NOT (#DiamondStep.S11)) AND "DB720_KuKa_MainCtrl".StatusIn.do_DiamondDetc_Pos) AND #Aux.DiamondDetcNOKTimer.Q 成立时，将 TRUE 传送到 "DB1148_PromptBeeper".Public.DiamondCoreNOK
   IF (((#DiamondStep.S9 AND NOT ("DB720_KuKa_MainCtrl".CmdOut.di_NotDectceDiamond)) AND NOT (#DiamondStep.S11)) AND "DB720_KuKa_MainCtrl".StatusIn.do_DiamondDetc_Pos) AND #Aux.DiamondDetcNOKTimer.Q THEN
       "DB1148_PromptBeeper".Public.DiamondCoreNOK := TRUE;
   END_IF;
   // 含义：将 (#DiamondStep.S9 AND #Aux.DiamondDetcOKTimer.Q) OR (#DiamondStep.S9 AND "DB720_KuKa_MainCtrl".CmdOut.di_NotDectceDiamond) OR (#DiamondStep.S9 AND #DiamondStep.S11) 赋给 #DiamondStep.S11
   #DiamondStep.S11 := (#DiamondStep.S9 AND #Aux.DiamondDetcOKTimer.Q) OR (#DiamondStep.S9 AND "DB720_KuKa_MainCtrl".CmdOut.di_NotDectceDiamond) OR (#DiamondStep.S9 AND #DiamondStep.S11);

   // ---------- 网络 12 ----------
   // 标题：水钻岩芯检测完成确认
   // 含义：条件 #DiamondStep.S11 AND NOT (#DiamondStep.S12) 成立时，将 TRUE 传送到 "DB720_KuKa_MainCtrl".CmdOut.di_DiamondDetc_Ack
   IF #DiamondStep.S11 AND NOT (#DiamondStep.S12) THEN
       "DB720_KuKa_MainCtrl".CmdOut.di_DiamondDetc_Ack := TRUE;
   END_IF;
   // 含义：将 ((#DiamondStep.S11 AND "DB720_KuKa_MainCtrl".StatusIn.do_Diamond_Don) AND "DB1080_Component".Robot.Status.HomePos) OR (#DiamondStep.S11 AND #DiamondStep.S12) 赋给 #DiamondStep.S12
   #DiamondStep.S12 := ((#DiamondStep.S11 AND "DB720_KuKa_MainCtrl".StatusIn.do_Diamond_Don) AND "DB1080_Component".Robot.Status.HomePos) OR (#DiamondStep.S11 AND #DiamondStep.S12);
   // 含义：将 ((#DiamondStep.S11 AND "DB720_KuKa_MainCtrl".StatusIn.do_Diamond_Don) AND "DB1080_Component".Robot.Status.HomePos) OR (#DiamondStep.S11 AND #DiamondStep.S12) 赋给 #DiamondStep.TaskDone
   #DiamondStep.TaskDone := ((#DiamondStep.S11 AND "DB720_KuKa_MainCtrl".StatusIn.do_Diamond_Don) AND "DB1080_Component".Robot.Status.HomePos) OR (#DiamondStep.S11 AND #DiamondStep.S12);

   // ---------- 网络 13 ----------
   // 含义：将 ((#DiamondStep.TaskDone OR #DiamondStep.ErrEnd OR #DiamondStep.ByPass OR #DiamondStep.S12) AND NOT (#DiamondStep.S13)) AND NOT (#DiamondStep.ErrEnd) 赋给 #DiamondStep.TaskIO
   #DiamondStep.TaskIO := ((#DiamondStep.TaskDone OR #DiamondStep.ErrEnd OR #DiamondStep.ByPass OR #DiamondStep.S12) AND NOT (#DiamondStep.S13)) AND NOT (#DiamondStep.ErrEnd);
   // 含义：将 ((#DiamondStep.TaskDone OR #DiamondStep.ErrEnd OR #DiamondStep.ByPass OR #DiamondStep.S12) AND NOT (#DiamondStep.S13)) AND #DiamondStep.ErrEnd 赋给 #DiamondStep.TaskNIO
   #DiamondStep.TaskNIO := ((#DiamondStep.TaskDone OR #DiamondStep.ErrEnd OR #DiamondStep.ByPass OR #DiamondStep.S12) AND NOT (#DiamondStep.S13)) AND #DiamondStep.ErrEnd;
   // 含义：条件 (#DiamondStep.TaskDone OR #DiamondStep.ErrEnd OR #DiamondStep.ByPass OR #DiamondStep.S12) AND NOT (#DiamondStep.S13) 成立时，将 FALSE 传送到 "DB720_KuKa_MainCtrl".CmdOut.di_DiamondDetc_Ack
   IF (#DiamondStep.TaskDone OR #DiamondStep.ErrEnd OR #DiamondStep.ByPass OR #DiamondStep.S12) AND NOT (#DiamondStep.S13) THEN
       "DB720_KuKa_MainCtrl".CmdOut.di_DiamondDetc_Ack := FALSE;
   END_IF;
   // 含义：将 #DiamondStep.TaskDone OR #DiamondStep.ErrEnd OR #DiamondStep.ByPass OR #DiamondStep.S12 赋给 #DiamondStep.S13
   #DiamondStep.S13 := #DiamondStep.TaskDone OR #DiamondStep.ErrEnd OR #DiamondStep.ByPass OR #DiamondStep.S12;

   // ---------- 网络 14 ----------
   // 含义：当 #DiamondStep.S13 为 TRUE 时置位 #DiamondStep.StepEnd，否则复位（触点→线圈）
   IF #DiamondStep.S13 THEN
       #DiamondStep.StepEnd := TRUE;
   ELSE
       #DiamondStep.StepEnd := FALSE;
   END_IF;

   // ---------- 网络 15 ----------
   // 含义：将 FALSE 赋给 #DiamondStep.StartCmd
   #DiamondStep.StartCmd := FALSE;

   // ---------- 网络 16 ----------
   // （空白网络）
END_FUNCTION_BLOCK

FUNCTION_BLOCK "FB1081_ValveCall"   // FB1081, SCL
{ S7_Optimized_Access := 'TRUE' }
// ============================================================
//  Block: FB1081_ValveCall
//  ============================================================
//  编号：FB1081
//  原始语言：LAD（规则翻译为 SCL）
//  含义：*****************************************************************************
//  *****************************************************************************
//  ***********************上海克来机电自动化工程有限公司************************
//  ***********************          V2014.10.25          ***********************
//  **********************                                 **********************
//  *****************************************************************************
//  *****************************************************************************
   VAR
      ST01 : Struct   // 静态变量
         Z01 : Struct   // 推力气缸
            ExtTPPB : Bool;   // 推力气缸
            RetTPPB : Bool;   // 推力气缸
            ExtPmt : Bool;   // 推力气缸
            RetPmt : Bool;   // 推力气缸
            IExtPos : Bool;   // 推力气缸
            IRetPos : Bool;   // 推力气缸
            TPSP1 : Bool;   // 推力气缸
            VentValveTPPB : Bool;   // 推力气缸
            ExtEVT : Bool;   // 推力气缸
            RetEVT : Bool;   // 推力气缸
            ExtPos : Bool;   // 推力气缸
            RetPos : Bool;   // 推力气缸
            ExtIng : Bool;   // 推力气缸
            RetIng : Bool;   // 推力气缸
            ExtErr : Bool;   // 推力气缸
            RetErr : Bool;   // 推力气缸
            ExtAuto : Bool;   // 推力气缸
            RetAuto : Bool;   // 推力气缸
            VentValveAuto : Bool;   // 推力气缸
            VentValve : Bool;   // 推力气缸
            Moving : Bool;   // 推力气缸
            RegTimer : Int;   // 推力气缸
         END_STRUCT;
         Z02 : Struct   // 辅助气缸
            ExtTPPB : Bool;   // 辅助气缸
            RetTPPB : Bool;   // 辅助气缸
            ExtPmt : Bool;   // 辅助气缸
            RetPmt : Bool;   // 辅助气缸
            IExtPos : Bool;   // 辅助气缸
            IRetPos : Bool;   // 辅助气缸
            TPSP1 : Bool;   // 辅助气缸
            VentValveTPPB : Bool;   // 辅助气缸
            ExtEVT : Bool;   // 辅助气缸
            RetEVT : Bool;   // 辅助气缸
            ExtPos : Bool;   // 辅助气缸
            RetPos : Bool;   // 辅助气缸
            ExtIng : Bool;   // 辅助气缸
            RetIng : Bool;   // 辅助气缸
            ExtErr : Bool;   // 辅助气缸
            RetErr : Bool;   // 辅助气缸
            ExtAuto : Bool;   // 辅助气缸
            RetAuto : Bool;   // 辅助气缸
            VentValveAuto : Bool;   // 辅助气缸
            VentValve : Bool;   // 辅助气缸
            Moving : Bool;   // 辅助气缸
            RegTimer : Int;   // 辅助气缸
         END_STRUCT;
         Z03 : Struct   // 左防尘盖夹紧缸
            ExtTPPB : Bool;   // 左防尘盖夹紧缸
            RetTPPB : Bool;   // 左防尘盖夹紧缸
            ExtPmt : Bool;   // 左防尘盖夹紧缸
            RetPmt : Bool;   // 左防尘盖夹紧缸
            IExtPos : Bool;   // 左防尘盖夹紧缸
            IRetPos : Bool;   // 左防尘盖夹紧缸
            TPSP1 : Bool;   // 左防尘盖夹紧缸
            VentValveTPPB : Bool;   // 左防尘盖夹紧缸
            ExtEVT : Bool;   // 左防尘盖夹紧缸
            RetEVT : Bool;   // 左防尘盖夹紧缸
            ExtPos : Bool;   // 左防尘盖夹紧缸
            RetPos : Bool;   // 左防尘盖夹紧缸
            ExtIng : Bool;   // 左防尘盖夹紧缸
            RetIng : Bool;   // 左防尘盖夹紧缸
            ExtErr : Bool;   // 左防尘盖夹紧缸
            RetErr : Bool;   // 左防尘盖夹紧缸
            ExtAuto : Bool;   // 左防尘盖夹紧缸
            RetAuto : Bool;   // 左防尘盖夹紧缸
            VentValveAuto : Bool;   // 左防尘盖夹紧缸
            VentValve : Bool;   // 左防尘盖夹紧缸
            Moving : Bool;   // 左防尘盖夹紧缸
            RegTimer : Int;   // 左防尘盖夹紧缸
         END_STRUCT;
         Z04 : Struct   // 右防尘盖夹紧缸
            ExtTPPB : Bool;   // 右防尘盖夹紧缸
            RetTPPB : Bool;   // 右防尘盖夹紧缸
            ExtPmt : Bool;   // 右防尘盖夹紧缸
            RetPmt : Bool;   // 右防尘盖夹紧缸
            IExtPos : Bool;   // 右防尘盖夹紧缸
            IRetPos : Bool;   // 右防尘盖夹紧缸
            TPSP1 : Bool;   // 右防尘盖夹紧缸
            VentValveTPPB : Bool;   // 右防尘盖夹紧缸
            ExtEVT : Bool;   // 右防尘盖夹紧缸
            RetEVT : Bool;   // 右防尘盖夹紧缸
            ExtPos : Bool;   // 右防尘盖夹紧缸
            RetPos : Bool;   // 右防尘盖夹紧缸
            ExtIng : Bool;   // 右防尘盖夹紧缸
            RetIng : Bool;   // 右防尘盖夹紧缸
            ExtErr : Bool;   // 右防尘盖夹紧缸
            RetErr : Bool;   // 右防尘盖夹紧缸
            ExtAuto : Bool;   // 右防尘盖夹紧缸
            RetAuto : Bool;   // 右防尘盖夹紧缸
            VentValveAuto : Bool;   // 右防尘盖夹紧缸
            VentValve : Bool;   // 右防尘盖夹紧缸
            Moving : Bool;   // 右防尘盖夹紧缸
            RegTimer : Int;   // 右防尘盖夹紧缸
         END_STRUCT;
         Z05 : Struct   // 枪电源
            ExtTPPB : Bool;   // 枪电源
            RetTPPB : Bool;   // 枪电源
            ExtPmt : Bool;   // 枪电源
            RetPmt : Bool;   // 枪电源
            IExtPos : Bool;   // 枪电源
            IRetPos : Bool;   // 枪电源
            TPSP1 : Bool;   // 枪电源
            VentValveTPPB : Bool;   // 枪电源
            ExtEVT : Bool;   // 枪电源
            RetEVT : Bool;   // 枪电源
            ExtPos : Bool;   // 枪电源
            RetPos : Bool;   // 枪电源
            ExtIng : Bool;   // 枪电源
            RetIng : Bool;   // 枪电源
            ExtErr : Bool;   // 枪电源
            RetErr : Bool;   // 枪电源
            ExtAuto : Bool;   // 枪电源
            RetAuto : Bool;   // 枪电源
            VentValveAuto : Bool;   // 枪电源
            VentValve : Bool;   // 枪电源
            Moving : Bool;   // 枪电源
            RegTimer : Int;   // 枪电源
         END_STRUCT;
         Z06 : Struct   // 摄像头防尘盖
            ExtTPPB : Bool;   // 水泥板吹气
            RetTPPB : Bool;   // 水泥板吹气
            ExtPmt : Bool;   // 水泥板吹气
            RetPmt : Bool;   // 水泥板吹气
            IExtPos : Bool;   // 水泥板吹气
            IRetPos : Bool;   // 水泥板吹气
            TPSP1 : Bool;   // 水泥板吹气
            VentValveTPPB : Bool;   // 水泥板吹气
            ExtEVT : Bool;   // 水泥板吹气
            RetEVT : Bool;   // 水泥板吹气
            ExtPos : Bool;   // 水泥板吹气
            RetPos : Bool;   // 水泥板吹气
            ExtIng : Bool;   // 水泥板吹气
            RetIng : Bool;   // 水泥板吹气
            ExtErr : Bool;   // 水泥板吹气
            RetErr : Bool;   // 水泥板吹气
            ExtAuto : Bool;   // 水泥板吹气
            RetAuto : Bool;   // 水泥板吹气
            VentValveAuto : Bool;   // 水泥板吹气
            VentValve : Bool;   // 水泥板吹气
            Moving : Bool;   // 水泥板吹气
            RegTimer : Int;   // 水泥板吹气
         END_STRUCT;
         Z07 : Struct   // 快换盘锁紧
            ExtTPPB : Bool;   // 快换盘锁紧
            RetTPPB : Bool;   // 快换盘锁紧
            ExtPmt : Bool;   // 快换盘锁紧
            RetPmt : Bool;   // 快换盘锁紧
            IExtPos : Bool;   // 快换盘锁紧
            IRetPos : Bool;   // 快换盘锁紧
            TPSP1 : Bool;   // 快换盘锁紧
            VentValveTPPB : Bool;   // 快换盘锁紧
            ExtEVT : Bool;   // 快换盘锁紧
            RetEVT : Bool;   // 快换盘锁紧
            ExtPos : Bool;   // 快换盘锁紧
            RetPos : Bool;   // 快换盘锁紧
            ExtIng : Bool;   // 快换盘锁紧
            RetIng : Bool;   // 快换盘锁紧
            ExtErr : Bool;   // 快换盘锁紧
            RetErr : Bool;   // 快换盘锁紧
            ExtAuto : Bool;   // 快换盘锁紧
            RetAuto : Bool;   // 快换盘解锁
            VentValveAuto : Bool;   // 快换盘锁紧
            VentValve : Bool;   // 快换盘锁紧
            Moving : Bool;   // 快换盘锁紧
            RegTimer : Int;   // 快换盘锁紧
         END_STRUCT;
         Z08 : Struct   // 参数写入
            ExtTPPB : Bool;   // 参数写入
            RetTPPB : Bool;   // 参数写入
            ExtPmt : Bool;   // 参数写入
            RetPmt : Bool;   // 参数写入
            IExtPos : Bool;   // 参数写入
            IRetPos : Bool;   // 参数写入
            TPSP1 : Bool;   // 参数写入
            VentValveTPPB : Bool;   // 参数写入
            ExtEVT : Bool;   // 参数写入
            RetEVT : Bool;   // 参数写入
            ExtPos : Bool;   // 参数写入
            RetPos : Bool;   // 参数写入
            ExtIng : Bool;   // 参数写入
            RetIng : Bool;   // 参数写入
            ExtErr : Bool;   // 参数写入
            RetErr : Bool;   // 参数写入
            ExtAuto : Bool;   // 参数写入
            RetAuto : Bool;   // 参数写入
            VentValveAuto : Bool;   // 参数写入
            VentValve : Bool;   // 参数写入
            Moving : Bool;   // 参数写入
            RegTimer : Int;   // 参数写入
         END_STRUCT;
         Z09 : Struct   // 凿击三爪卡盘夹爪气缸
            ExtTPPB : Bool := FALSE;   // 凿击三爪卡盘夹爪气缸
            RetTPPB : Bool := FALSE;   // 凿击三爪卡盘夹爪气缸
            ExtPmt : Bool := FALSE;   // 凿击三爪卡盘夹爪气缸
            RetPmt : Bool := FALSE;   // 凿击三爪卡盘夹爪气缸
            IExtPos : Bool := FALSE;   // 凿击三爪卡盘夹爪气缸
            IRetPos : Bool := FALSE;   // 凿击三爪卡盘夹爪气缸
            TPSP1 : Bool := FALSE;   // 凿击三爪卡盘夹爪气缸
            VentValveTPPB : Bool := FALSE;   // 凿击三爪卡盘夹爪气缸
            ExtEVT : Bool := FALSE;   // 凿击三爪卡盘夹爪气缸
            RetEVT : Bool := FALSE;   // 凿击三爪卡盘夹爪气缸
            ExtPos : Bool := FALSE;   // 凿击三爪卡盘夹爪气缸
            RetPos : Bool := FALSE;   // 凿击三爪卡盘夹爪气缸
            ExtIng : Bool := FALSE;   // 凿击三爪卡盘夹爪气缸
            RetIng : Bool := FALSE;   // 凿击三爪卡盘夹爪气缸
            ExtErr : Bool := FALSE;   // 凿击三爪卡盘夹爪气缸
            RetErr : Bool := FALSE;   // 凿击三爪卡盘夹爪气缸
            ExtAuto : Bool := FALSE;   // 凿击三爪卡盘夹爪气缸
            RetAuto : Bool := FALSE;   // 凿击三爪卡盘夹爪气缸
            VentValveAuto : Bool := FALSE;   // 凿击三爪卡盘夹爪气缸
            VentValve : Bool := FALSE;   // 凿击三爪卡盘夹爪气缸
            Moving : Bool := FALSE;   // 凿击三爪卡盘夹爪气缸
            RegTimer : Int := 0;   // 凿击三爪卡盘夹爪气缸
         END_STRUCT;
      END_STRUCT;
      "Time" : Struct   // 静态变量
         ST01Z03EXT : IEC_TIMER;   // Z03.A工位防尘罩伸出延时
         ST01Z03RetT : IEC_TIMER;   // Z03.A工位防尘罩缩回延时
         ST01Z04EXT : IEC_TIMER;   // Z04.B工位防尘罩伸出延时
         ST01Z04RET : IEC_TIMER;   // Z04.B工位防尘罩缩回延时
         ST01Z07EXT : IEC_TIMER;   // Z07.快换盘伸出延时
         ST01Z07RET : IEC_TIMER;   // Z07.快换盘缩回延时
         ST01Z08EXT : IEC_TIMER;   // Z08.参数写入伸出延时
         ST01Z08RET : IEC_TIMER;   // Z08.参数写入缩回延时
         ST01Z09EXT : IEC_TIMER;   // Z09.三爪卡盘气缸伸出延时
      END_STRUCT;
      EdgeDetc : Struct   // 静态变量
         Pulse : Array[0..15] of Bool;   // 静态变量
      END_STRUCT;
      PT : Time;   // 静态变量
      ET : Time;   // 静态变量
      IN : Bool;   // 静态变量
      Q : Bool;   // 静态变量
   END_VAR
   VAR_TEMP
      OverAllPmt : Bool;   // 临时变量
   END_VAR
BEGIN

   // ---------- 网络 1 ----------
   // 标题：ModeSwitch模式开关
   // 含义：当 "DB1001_SysMode".SubSysMode.Mode.ManMode 为 TRUE 时置位 "DB1200_FB_std_Switch".ManMode，否则复位（触点→线圈）
   IF "DB1001_SysMode".SubSysMode.Mode.ManMode THEN
       "DB1200_FB_std_Switch".ManMode := TRUE;
   ELSE
       "DB1200_FB_std_Switch".ManMode := FALSE;
   END_IF;
   // 含义：当 "DB1001_SysMode".SubSysMode.Mode.AllMode 为 TRUE 时置位 "DB1200_FB_std_Switch".AllMode，否则复位（触点→线圈）
   IF "DB1001_SysMode".SubSysMode.Mode.AllMode THEN
       "DB1200_FB_std_Switch".AllMode := TRUE;
   ELSE
       "DB1200_FB_std_Switch".AllMode := FALSE;
   END_IF;
   // 含义：当 "DB1001_SysMode".SubSysMode.Mode.EMMode 为 TRUE 时置位 "DB1200_FB_std_Switch".EMMode，否则复位（触点→线圈）
   IF "DB1001_SysMode".SubSysMode.Mode.EMMode THEN
       "DB1200_FB_std_Switch".EMMode := TRUE;
   ELSE
       "DB1200_FB_std_Switch".EMMode := FALSE;
   END_IF;
   // 含义：条件 "DB1001_SysMode".SubSysMode.Mode.EMMode 成立时，将 TRUE 传送到 #ST01.Z07.RetAuto
   IF "DB1001_SysMode".SubSysMode.Mode.EMMode THEN
       #ST01.Z07.RetAuto := TRUE;
   END_IF;
   // 含义：将 FALSE 赋给 "DB1200_FB_std_Switch".OprNotPmt
   "DB1200_FB_std_Switch".OprNotPmt := FALSE;
   // 含义：将 ("DB1001_SysMode".SubSysMode.Mode.AllMode AND NOT ("DB1080_Component".SafetyDoor.i_DoorOverRide)) AND "ICurtainsOK" 赋给 #OverAllPmt
   #OverAllPmt := ("DB1001_SysMode".SubSysMode.Mode.AllMode AND NOT ("DB1080_Component".SafetyDoor.i_DoorOverRide)) AND "ICurtainsOK";

   // ---------- 网络 2 ----------
   // 标题：Z01--->推力气缸
   // 含义：当 "IZ02RetPos" 为 TRUE 时置位 #ST01.Z01.IRetPos，否则复位（触点→线圈）
   IF "IZ02RetPos" THEN
       #ST01.Z01.IRetPos := TRUE;
   ELSE
       #ST01.Z01.IRetPos := FALSE;
   END_IF;
   // 含义：当 #ST01.Z01.ExtEVT 为 TRUE 时置位 #ST01.Z01.IExtPos，否则复位（触点→线圈）
   IF #ST01.Z01.ExtEVT THEN
       #ST01.Z01.IExtPos := TRUE;
   ELSE
       #ST01.Z01.IExtPos := FALSE;
   END_IF;
   // 含义：将 (NOT (#ST01.Z01.ExtEVT) AND #ST01.Z01.IRetPos) AND NOT (#ST01.Z01.IExtPos) 赋给 #ST01.Z01.RetPos
   #ST01.Z01.RetPos := (NOT (#ST01.Z01.ExtEVT) AND #ST01.Z01.IRetPos) AND NOT (#ST01.Z01.IExtPos);
   // 含义：将 (NOT (#ST01.Z01.ExtEVT) AND #ST01.Z01.IRetPos) AND NOT (#ST01.Z01.IExtPos) 赋给 "DB1900_Communication_PC".Send.Z01RetPos
   "DB1900_Communication_PC".Send.Z01RetPos := (NOT (#ST01.Z01.ExtEVT) AND #ST01.Z01.IRetPos) AND NOT (#ST01.Z01.IExtPos);
   // 含义：将 (NOT (#ST01.Z01.RetEVT) AND NOT (#ST01.Z01.IRetPos)) AND #ST01.Z01.IExtPos 赋给 #ST01.Z01.ExtPos
   #ST01.Z01.ExtPos := (NOT (#ST01.Z01.RetEVT) AND NOT (#ST01.Z01.IRetPos)) AND #ST01.Z01.IExtPos;
   // 含义：将 (NOT (#ST01.Z01.RetEVT) AND NOT (#ST01.Z01.IRetPos)) AND #ST01.Z01.IExtPos 赋给 "DB1900_Communication_PC".Send.Z01ExtPos
   "DB1900_Communication_PC".Send.Z01ExtPos := (NOT (#ST01.Z01.RetEVT) AND NOT (#ST01.Z01.IRetPos)) AND #ST01.Z01.IExtPos;
   // 含义：当 #OverAllPmt 为 TRUE 时置位 #ST01.Z01.ExtPmt，否则复位（触点→线圈）
   IF #OverAllPmt THEN
       #ST01.Z01.ExtPmt := TRUE;
   ELSE
       #ST01.Z01.ExtPmt := FALSE;
   END_IF;
   // 含义：当 #OverAllPmt 为 TRUE 时置位 #ST01.Z01.RetPmt，否则复位（触点→线圈）
   IF #OverAllPmt THEN
       #ST01.Z01.RetPmt := TRUE;
   ELSE
       #ST01.Z01.RetPmt := FALSE;
   END_IF;
   // 含义：调用块/实例 "DB1200_FB_std_Switch"，参数：CylinderCmd := #ST01.Z01
   "DB1200_FB_std_Switch"(CylinderCmd := #ST01.Z01);
   // 含义：当 #ST01.Z01.ExtIng 为 TRUE 时置位 "DB1146_PromptFree".ST01.Z01ExtIng，否则复位（触点→线圈）
   IF #ST01.Z01.ExtIng THEN
       "DB1146_PromptFree".ST01.Z01ExtIng := TRUE;
   ELSE
       "DB1146_PromptFree".ST01.Z01ExtIng := FALSE;
   END_IF;
   // 含义：当 #ST01.Z01.RetIng 为 TRUE 时置位 "DB1146_PromptFree".ST01.Z01RetIng，否则复位（触点→线圈）
   IF #ST01.Z01.RetIng THEN
       "DB1146_PromptFree".ST01.Z01RetIng := TRUE;
   ELSE
       "DB1146_PromptFree".ST01.Z01RetIng := FALSE;
   END_IF;
   // 含义：当 #ST01.Z01.ExtErr 为 TRUE 时置位 "DB1148_PromptBeeper".ST01.Z01ExtErr，否则复位（触点→线圈）
   IF #ST01.Z01.ExtErr THEN
       "DB1148_PromptBeeper".ST01.Z01ExtErr := TRUE;
   ELSE
       "DB1148_PromptBeeper".ST01.Z01ExtErr := FALSE;
   END_IF;
   // 含义：当 #ST01.Z01.RetErr 为 TRUE 时置位 "DB1148_PromptBeeper".ST01.Z01RetErr，否则复位（触点→线圈）
   IF #ST01.Z01.RetErr THEN
       "DB1148_PromptBeeper".ST01.Z01RetErr := TRUE;
   ELSE
       "DB1148_PromptBeeper".ST01.Z01RetErr := FALSE;
   END_IF;
   // 含义：将 #ST01.Z01.ExtEVT AND NOT ("DB1148_PromptBeeper".Public.AirPressureLow) 赋给 "QZ01ExtEvt"
   "QZ01ExtEvt" := #ST01.Z01.ExtEVT AND NOT ("DB1148_PromptBeeper".Public.AirPressureLow);
   // 含义：将 #ST01.Z01.RetEVT AND NOT ("DB1148_PromptBeeper".Public.AirPressureLow) 赋给 "QZ01RetEvt"
   "QZ01RetEvt" := #ST01.Z01.RetEVT AND NOT ("DB1148_PromptBeeper".Public.AirPressureLow);
   // 含义：条件 "ManMode_M" AND "DB1900_Communication_PC".Recv.Z01ExtTPPB 成立时，将 TRUE 传送到 #ST01.Z01.ExtAuto
   IF "ManMode_M" AND "DB1900_Communication_PC".Recv.Z01ExtTPPB THEN
       #ST01.Z01.ExtAuto := TRUE;
   END_IF;
   // 含义：条件 "ManMode_M" AND "DB1900_Communication_PC".Recv.Z01RetTPPB 成立时，将 TRUE 传送到 #ST01.Z01.RetAuto
   IF "ManMode_M" AND "DB1900_Communication_PC".Recv.Z01RetTPPB THEN
       #ST01.Z01.RetAuto := TRUE;
   END_IF;
   // 含义：条件 "ManMode_M" AND "DB1900_Communication_PC".Recv.Z01VentValveTPPB 成立时，将 TRUE 传送到 #ST01.Z01.VentValveAuto
   IF "ManMode_M" AND "DB1900_Communication_PC".Recv.Z01VentValveTPPB THEN
       #ST01.Z01.VentValveAuto := TRUE;
   END_IF;
   // 含义：条件 "ManMode_M" AND "DB1900_Communication_PC".Recv.Z02VentValveTPPB 成立时，将 TRUE 传送到 #ST01.Z02.VentValveAuto
   IF "ManMode_M" AND "DB1900_Communication_PC".Recv.Z02VentValveTPPB THEN
       #ST01.Z02.VentValveAuto := TRUE;
   END_IF;
   // 含义：将 "ManMode_M" AND #ST01.Z01.VentValve 赋给 "DB1900_Communication_PC".Send.Z01VentValve
   "DB1900_Communication_PC".Send.Z01VentValve := "ManMode_M" AND #ST01.Z01.VentValve;
   // 含义：将 "ManMode_M" AND #ST01.Z02.VentValve 赋给 "DB1900_Communication_PC".Send.Z02VentValve
   "DB1900_Communication_PC".Send.Z02VentValve := "ManMode_M" AND #ST01.Z02.VentValve;

   // ---------- 网络 3 ----------
   // 标题：Z02--->辅助气缸
   // 含义：当 #ST01.Z02.RetEVT 为 TRUE 时置位 #ST01.Z02.IRetPos，否则复位（触点→线圈）
   IF #ST01.Z02.RetEVT THEN
       #ST01.Z02.IRetPos := TRUE;
   ELSE
       #ST01.Z02.IRetPos := FALSE;
   END_IF;
   // 含义：当 #ST01.Z02.ExtEVT 为 TRUE 时置位 #ST01.Z02.IExtPos，否则复位（触点→线圈）
   IF #ST01.Z02.ExtEVT THEN
       #ST01.Z02.IExtPos := TRUE;
   ELSE
       #ST01.Z02.IExtPos := FALSE;
   END_IF;
   // 含义：将 (NOT (#ST01.Z02.ExtEVT) AND #ST01.Z02.IRetPos) AND NOT (#ST01.Z02.IExtPos) 赋给 #ST01.Z02.RetPos
   #ST01.Z02.RetPos := (NOT (#ST01.Z02.ExtEVT) AND #ST01.Z02.IRetPos) AND NOT (#ST01.Z02.IExtPos);
   // 含义：将 (NOT (#ST01.Z02.ExtEVT) AND #ST01.Z02.IRetPos) AND NOT (#ST01.Z02.IExtPos) 赋给 "DB1900_Communication_PC".Send.Z02RetPos
   "DB1900_Communication_PC".Send.Z02RetPos := (NOT (#ST01.Z02.ExtEVT) AND #ST01.Z02.IRetPos) AND NOT (#ST01.Z02.IExtPos);
   // 含义：将 (NOT (#ST01.Z02.RetEVT) AND NOT (#ST01.Z02.IRetPos)) AND #ST01.Z02.IExtPos 赋给 #ST01.Z02.ExtPos
   #ST01.Z02.ExtPos := (NOT (#ST01.Z02.RetEVT) AND NOT (#ST01.Z02.IRetPos)) AND #ST01.Z02.IExtPos;
   // 含义：将 (NOT (#ST01.Z02.RetEVT) AND NOT (#ST01.Z02.IRetPos)) AND #ST01.Z02.IExtPos 赋给 "DB1900_Communication_PC".Send.Z02ExtPos
   "DB1900_Communication_PC".Send.Z02ExtPos := (NOT (#ST01.Z02.RetEVT) AND NOT (#ST01.Z02.IRetPos)) AND #ST01.Z02.IExtPos;
   // 含义：当 #OverAllPmt 为 TRUE 时置位 #ST01.Z02.ExtPmt，否则复位（触点→线圈）
   IF #OverAllPmt THEN
       #ST01.Z02.ExtPmt := TRUE;
   ELSE
       #ST01.Z02.ExtPmt := FALSE;
   END_IF;
   // 含义：当 #OverAllPmt 为 TRUE 时置位 #ST01.Z02.RetPmt，否则复位（触点→线圈）
   IF #OverAllPmt THEN
       #ST01.Z02.RetPmt := TRUE;
   ELSE
       #ST01.Z02.RetPmt := FALSE;
   END_IF;
   // 含义：调用块/实例 "DB1200_FB_std_Switch"，参数：CylinderCmd := #ST01.Z02
   "DB1200_FB_std_Switch"(CylinderCmd := #ST01.Z02);
   // 含义：当 #ST01.Z02.ExtIng 为 TRUE 时置位 "DB1146_PromptFree".ST01.Z02ExtIng，否则复位（触点→线圈）
   IF #ST01.Z02.ExtIng THEN
       "DB1146_PromptFree".ST01.Z02ExtIng := TRUE;
   ELSE
       "DB1146_PromptFree".ST01.Z02ExtIng := FALSE;
   END_IF;
   // 含义：当 #ST01.Z02.RetIng 为 TRUE 时置位 "DB1146_PromptFree".ST01.Z02RetIng，否则复位（触点→线圈）
   IF #ST01.Z02.RetIng THEN
       "DB1146_PromptFree".ST01.Z02RetIng := TRUE;
   ELSE
       "DB1146_PromptFree".ST01.Z02RetIng := FALSE;
   END_IF;
   // 含义：当 #ST01.Z02.ExtErr 为 TRUE 时置位 "DB1148_PromptBeeper".ST01.Z02ExtErr，否则复位（触点→线圈）
   IF #ST01.Z02.ExtErr THEN
       "DB1148_PromptBeeper".ST01.Z02ExtErr := TRUE;
   ELSE
       "DB1148_PromptBeeper".ST01.Z02ExtErr := FALSE;
   END_IF;
   // 含义：当 #ST01.Z02.RetErr 为 TRUE 时置位 "DB1148_PromptBeeper".ST01.Z02RetErr，否则复位（触点→线圈）
   IF #ST01.Z02.RetErr THEN
       "DB1148_PromptBeeper".ST01.Z02RetErr := TRUE;
   ELSE
       "DB1148_PromptBeeper".ST01.Z02RetErr := FALSE;
   END_IF;
   // 含义：将 #ST01.Z02.ExtEVT AND NOT ("DB1148_PromptBeeper".Public.AirPressureLow) 赋给 "QZ02ExtEvt"
   "QZ02ExtEvt" := #ST01.Z02.ExtEVT AND NOT ("DB1148_PromptBeeper".Public.AirPressureLow);
   // 含义：将 #ST01.Z02.RetEVT AND NOT ("DB1148_PromptBeeper".Public.AirPressureLow) 赋给 "QZ02RetEvt"
   "QZ02RetEvt" := #ST01.Z02.RetEVT AND NOT ("DB1148_PromptBeeper".Public.AirPressureLow);
   // 含义：条件 "ManMode_M" AND "DB1900_Communication_PC".Recv.Z02ExtTPPB 成立时，将 TRUE 传送到 #ST01.Z02.ExtAuto
   IF "ManMode_M" AND "DB1900_Communication_PC".Recv.Z02ExtTPPB THEN
       #ST01.Z02.ExtAuto := TRUE;
   END_IF;
   // 含义：条件 "ManMode_M" AND "DB1900_Communication_PC".Recv.Z02RetTPPB 成立时，将 TRUE 传送到 #ST01.Z02.RetAuto
   IF "ManMode_M" AND "DB1900_Communication_PC".Recv.Z02RetTPPB THEN
       #ST01.Z02.RetAuto := TRUE;
   END_IF;

   // ---------- 网络 4 ----------
   // 标题：Z03--->A工位防尘盖夹紧缸
   // 含义：当 "AStation_IZ03RetPos" 为 TRUE 时置位 #ST01.Z03.IRetPos，否则复位（触点→线圈）
   IF "AStation_IZ03RetPos" THEN
       #ST01.Z03.IRetPos := TRUE;
   ELSE
       #ST01.Z03.IRetPos := FALSE;
   END_IF;
   // 含义：当 "AStation_IZ03ExtPos" 为 TRUE 时置位 #ST01.Z03.IExtPos，否则复位（触点→线圈）
   IF "AStation_IZ03ExtPos" THEN
       #ST01.Z03.IExtPos := TRUE;
   ELSE
       #ST01.Z03.IExtPos := FALSE;
   END_IF;
   // 含义：将 (NOT (#ST01.Z03.ExtEVT) AND #ST01.Z03.IRetPos) AND NOT (#ST01.Z03.IExtPos) 赋给 #ST01.Z03.RetPos
   #ST01.Z03.RetPos := (NOT (#ST01.Z03.ExtEVT) AND #ST01.Z03.IRetPos) AND NOT (#ST01.Z03.IExtPos);
   // 含义：将 (NOT (#ST01.Z03.ExtEVT) AND #ST01.Z03.IRetPos) AND NOT (#ST01.Z03.IExtPos) 赋给 "DB1900_Communication_PC".Send.Z03RetPos
   "DB1900_Communication_PC".Send.Z03RetPos := (NOT (#ST01.Z03.ExtEVT) AND #ST01.Z03.IRetPos) AND NOT (#ST01.Z03.IExtPos);
   // 含义：将 (NOT (#ST01.Z03.RetEVT) AND NOT (#ST01.Z03.IRetPos)) AND #ST01.Z03.IExtPos 赋给 #ST01.Z03.ExtPos
   #ST01.Z03.ExtPos := (NOT (#ST01.Z03.RetEVT) AND NOT (#ST01.Z03.IRetPos)) AND #ST01.Z03.IExtPos;
   // 含义：将 (NOT (#ST01.Z03.RetEVT) AND NOT (#ST01.Z03.IRetPos)) AND #ST01.Z03.IExtPos 赋给 "DB1900_Communication_PC".Send.Z03ExtPos
   "DB1900_Communication_PC".Send.Z03ExtPos := (NOT (#ST01.Z03.RetEVT) AND NOT (#ST01.Z03.IRetPos)) AND #ST01.Z03.IExtPos;
   // 含义：当 #OverAllPmt 为 TRUE 时置位 #ST01.Z03.ExtPmt，否则复位（触点→线圈）
   IF #OverAllPmt THEN
       #ST01.Z03.ExtPmt := TRUE;
   ELSE
       #ST01.Z03.ExtPmt := FALSE;
   END_IF;
   // 含义：当 #OverAllPmt 为 TRUE 时置位 #ST01.Z03.RetPmt，否则复位（触点→线圈）
   IF #OverAllPmt THEN
       #ST01.Z03.RetPmt := TRUE;
   ELSE
       #ST01.Z03.RetPmt := FALSE;
   END_IF;
   // 含义：调用块/实例 "DB1200_FB_std_Switch"，参数：CylinderCmd := #ST01.Z03
   "DB1200_FB_std_Switch"(CylinderCmd := #ST01.Z03);
   // 含义：当 #ST01.Z03.ExtIng 为 TRUE 时置位 "DB1146_PromptFree".ST01.Z03ExtIng，否则复位（触点→线圈）
   IF #ST01.Z03.ExtIng THEN
       "DB1146_PromptFree".ST01.Z03ExtIng := TRUE;
   ELSE
       "DB1146_PromptFree".ST01.Z03ExtIng := FALSE;
   END_IF;
   // 含义：当 #ST01.Z03.RetIng 为 TRUE 时置位 "DB1146_PromptFree".ST01.Z03RetIng，否则复位（触点→线圈）
   IF #ST01.Z03.RetIng THEN
       "DB1146_PromptFree".ST01.Z03RetIng := TRUE;
   ELSE
       "DB1146_PromptFree".ST01.Z03RetIng := FALSE;
   END_IF;
   // 含义：将 #ST01.Z03.ExtErr AND #Time.ST01Z03EXT.Q 赋给 "DB1148_PromptBeeper".ST01.Z03ExtErr
   "DB1148_PromptBeeper".ST01.Z03ExtErr := #ST01.Z03.ExtErr AND #Time.ST01Z03EXT.Q;
   // 含义：调用定时器实例 #Time.ST01Z03EXT.TON
   #Time.ST01Z03EXT.TON(IN := #ST01.Z03.ExtErr,
                        PT := T#6s);
   // 含义：将 #ST01.Z03.RetErr AND #Time.ST01Z03RetT.Q 赋给 "DB1148_PromptBeeper".ST01.Z03RetErr
   "DB1148_PromptBeeper".ST01.Z03RetErr := #ST01.Z03.RetErr AND #Time.ST01Z03RetT.Q;
   // 含义：调用定时器实例 #Time.ST01Z03RetT.TON
   #Time.ST01Z03RetT.TON(IN := #ST01.Z03.RetErr,
                         PT := T#6s);
   // 含义：当 #ST01.Z03.ExtEVT 为 TRUE 时置位 "QZ03ExtEvt"，否则复位（触点→线圈）
   IF #ST01.Z03.ExtEVT THEN
       "QZ03ExtEvt" := TRUE;
   ELSE
       "QZ03ExtEvt" := FALSE;
   END_IF;
   // 含义：当 #ST01.Z03.RetEVT 为 TRUE 时置位 "QZ03RetEvt"，否则复位（触点→线圈）
   IF #ST01.Z03.RetEVT THEN
       "QZ03RetEvt" := TRUE;
   ELSE
       "QZ03RetEvt" := FALSE;
   END_IF;
   // 含义：条件 "ManMode_M" AND "DB1900_Communication_PC".Recv.Z03ExtTPPB 成立时，将 TRUE 传送到 #ST01.Z03.ExtAuto
   IF "ManMode_M" AND "DB1900_Communication_PC".Recv.Z03ExtTPPB THEN
       #ST01.Z03.ExtAuto := TRUE;
   END_IF;
   // 含义：条件 "ManMode_M" AND "DB1900_Communication_PC".Recv.Z03RetTPPB 成立时，将 TRUE 传送到 #ST01.Z03.RetAuto
   IF "ManMode_M" AND "DB1900_Communication_PC".Recv.Z03RetTPPB THEN
       #ST01.Z03.RetAuto := TRUE;
   END_IF;

   // ---------- 网络 5 ----------
   // 标题：Z04--->B工位防尘盖夹紧缸
   // 含义：当 "BStation_IZ04RetPos" 为 TRUE 时置位 #ST01.Z04.IRetPos，否则复位（触点→线圈）
   IF "BStation_IZ04RetPos" THEN
       #ST01.Z04.IRetPos := TRUE;
   ELSE
       #ST01.Z04.IRetPos := FALSE;
   END_IF;
   // 含义：当 "BStation_IZ04ExtPos" 为 TRUE 时置位 #ST01.Z04.IExtPos，否则复位（触点→线圈）
   IF "BStation_IZ04ExtPos" THEN
       #ST01.Z04.IExtPos := TRUE;
   ELSE
       #ST01.Z04.IExtPos := FALSE;
   END_IF;
   // 含义：将 (NOT (#ST01.Z04.ExtEVT) AND #ST01.Z04.IRetPos) AND NOT (#ST01.Z04.IExtPos) 赋给 #ST01.Z04.RetPos
   #ST01.Z04.RetPos := (NOT (#ST01.Z04.ExtEVT) AND #ST01.Z04.IRetPos) AND NOT (#ST01.Z04.IExtPos);
   // 含义：将 (NOT (#ST01.Z04.ExtEVT) AND #ST01.Z04.IRetPos) AND NOT (#ST01.Z04.IExtPos) 赋给 "DB1900_Communication_PC".Send.Z04RetPos
   "DB1900_Communication_PC".Send.Z04RetPos := (NOT (#ST01.Z04.ExtEVT) AND #ST01.Z04.IRetPos) AND NOT (#ST01.Z04.IExtPos);
   // 含义：将 (NOT (#ST01.Z04.RetEVT) AND NOT (#ST01.Z04.IRetPos)) AND #ST01.Z04.IExtPos 赋给 #ST01.Z04.ExtPos
   #ST01.Z04.ExtPos := (NOT (#ST01.Z04.RetEVT) AND NOT (#ST01.Z04.IRetPos)) AND #ST01.Z04.IExtPos;
   // 含义：将 (NOT (#ST01.Z04.RetEVT) AND NOT (#ST01.Z04.IRetPos)) AND #ST01.Z04.IExtPos 赋给 "DB1900_Communication_PC".Send.Z04ExtPos
   "DB1900_Communication_PC".Send.Z04ExtPos := (NOT (#ST01.Z04.RetEVT) AND NOT (#ST01.Z04.IRetPos)) AND #ST01.Z04.IExtPos;
   // 含义：当 #OverAllPmt 为 TRUE 时置位 #ST01.Z04.ExtPmt，否则复位（触点→线圈）
   IF #OverAllPmt THEN
       #ST01.Z04.ExtPmt := TRUE;
   ELSE
       #ST01.Z04.ExtPmt := FALSE;
   END_IF;
   // 含义：当 #OverAllPmt 为 TRUE 时置位 #ST01.Z04.RetPmt，否则复位（触点→线圈）
   IF #OverAllPmt THEN
       #ST01.Z04.RetPmt := TRUE;
   ELSE
       #ST01.Z04.RetPmt := FALSE;
   END_IF;
   // 含义：调用块/实例 "DB1200_FB_std_Switch"，参数：CylinderCmd := #ST01.Z04
   "DB1200_FB_std_Switch"(CylinderCmd := #ST01.Z04);
   // 含义：当 #ST01.Z04.ExtIng 为 TRUE 时置位 "DB1146_PromptFree".ST01.Z04ExtIng，否则复位（触点→线圈）
   IF #ST01.Z04.ExtIng THEN
       "DB1146_PromptFree".ST01.Z04ExtIng := TRUE;
   ELSE
       "DB1146_PromptFree".ST01.Z04ExtIng := FALSE;
   END_IF;
   // 含义：当 #ST01.Z04.RetIng 为 TRUE 时置位 "DB1146_PromptFree".ST01.Z04RetIng，否则复位（触点→线圈）
   IF #ST01.Z04.RetIng THEN
       "DB1146_PromptFree".ST01.Z04RetIng := TRUE;
   ELSE
       "DB1146_PromptFree".ST01.Z04RetIng := FALSE;
   END_IF;
   // 含义：将 #ST01.Z04.ExtErr AND #Time.ST01Z04EXT.Q 赋给 "DB1148_PromptBeeper".ST01.Z04ExtErr
   "DB1148_PromptBeeper".ST01.Z04ExtErr := #ST01.Z04.ExtErr AND #Time.ST01Z04EXT.Q;
   // 含义：调用定时器实例 #Time.ST01Z04EXT.TON
   #Time.ST01Z04EXT.TON(IN := #ST01.Z04.ExtErr,
                        PT := T#4s);
   // 含义：将 #ST01.Z04.RetErr AND #Time.ST01Z04RET.Q 赋给 "DB1148_PromptBeeper".ST01.Z04RetErr
   "DB1148_PromptBeeper".ST01.Z04RetErr := #ST01.Z04.RetErr AND #Time.ST01Z04RET.Q;
   // 含义：调用定时器实例 #Time.ST01Z04RET.TON
   #Time.ST01Z04RET.TON(IN := #ST01.Z04.RetErr,
                        PT := T#4s);
   // 含义：当 #ST01.Z04.ExtEVT 为 TRUE 时置位 "QZ04ExtEvt"，否则复位（触点→线圈）
   IF #ST01.Z04.ExtEVT THEN
       "QZ04ExtEvt" := TRUE;
   ELSE
       "QZ04ExtEvt" := FALSE;
   END_IF;
   // 含义：当 #ST01.Z04.RetEVT 为 TRUE 时置位 "QZ04RetEvt"，否则复位（触点→线圈）
   IF #ST01.Z04.RetEVT THEN
       "QZ04RetEvt" := TRUE;
   ELSE
       "QZ04RetEvt" := FALSE;
   END_IF;
   // 含义：条件 "ManMode_M" AND "DB1900_Communication_PC".Recv.Z04ExtTPPB 成立时，将 TRUE 传送到 #ST01.Z04.ExtAuto
   IF "ManMode_M" AND "DB1900_Communication_PC".Recv.Z04ExtTPPB THEN
       #ST01.Z04.ExtAuto := TRUE;
   END_IF;
   // 含义：条件 "ManMode_M" AND "DB1900_Communication_PC".Recv.Z04RetTPPB 成立时，将 TRUE 传送到 #ST01.Z04.RetAuto
   IF "ManMode_M" AND "DB1900_Communication_PC".Recv.Z04RetTPPB THEN
       #ST01.Z04.RetAuto := TRUE;
   END_IF;

   // ---------- 网络 6 ----------
   // 标题：Z05--->枪电源
   // 注释：必须上位机先打开电源箱，PLC才能控制气缸接通,  三爪卡盘复用为电源开关控制气缸
   // 含义：当 "DB1900_Communication_PC".Recv.Z05RetTPPB 为 TRUE 时置位 #ST01.Z05.IRetPos，否则复位（触点→线圈）
   IF "DB1900_Communication_PC".Recv.Z05RetTPPB THEN
       #ST01.Z05.IRetPos := TRUE;
   ELSE
       #ST01.Z05.IRetPos := FALSE;
   END_IF;
   // 含义：当 "DB1900_Communication_PC".Recv.Z05ExtTPPB 为 TRUE 时置位 #ST01.Z05.IExtPos，否则复位（触点→线圈）
   IF "DB1900_Communication_PC".Recv.Z05ExtTPPB THEN
       #ST01.Z05.IExtPos := TRUE;
   ELSE
       #ST01.Z05.IExtPos := FALSE;
   END_IF;
   // 含义：将 #ST01.Z05.IRetPos AND NOT (#ST01.Z05.IExtPos) 赋给 #ST01.Z05.RetPos
   #ST01.Z05.RetPos := #ST01.Z05.IRetPos AND NOT (#ST01.Z05.IExtPos);
   // 含义：将 NOT (#ST01.Z05.IRetPos) AND #ST01.Z05.IExtPos 赋给 #ST01.Z05.ExtPos
   #ST01.Z05.ExtPos := NOT (#ST01.Z05.IRetPos) AND #ST01.Z05.IExtPos;
   // 含义：当 #OverAllPmt 为 TRUE 时置位 #ST01.Z05.ExtPmt，否则复位（触点→线圈）
   IF #OverAllPmt THEN
       #ST01.Z05.ExtPmt := TRUE;
   ELSE
       #ST01.Z05.ExtPmt := FALSE;
   END_IF;
   // 含义：当 #OverAllPmt 为 TRUE 时置位 #ST01.Z05.RetPmt，否则复位（触点→线圈）
   IF #OverAllPmt THEN
       #ST01.Z05.RetPmt := TRUE;
   ELSE
       #ST01.Z05.RetPmt := FALSE;
   END_IF;
   // 含义：调用块/实例 "DB1200_FB_std_Switch"，参数：CylinderCmd := #ST01.Z05
   "DB1200_FB_std_Switch"(CylinderCmd := #ST01.Z05);
   // 含义：当 #ST01.Z05.ExtIng 为 TRUE 时置位 "DB1146_PromptFree".ST01.Z05ExtIng，否则复位（触点→线圈）
   IF #ST01.Z05.ExtIng THEN
       "DB1146_PromptFree".ST01.Z05ExtIng := TRUE;
   ELSE
       "DB1146_PromptFree".ST01.Z05ExtIng := FALSE;
   END_IF;
   // 含义：当 #ST01.Z05.RetIng 为 TRUE 时置位 "DB1146_PromptFree".ST01.Z05RetIng，否则复位（触点→线圈）
   IF #ST01.Z05.RetIng THEN
       "DB1146_PromptFree".ST01.Z05RetIng := TRUE;
   ELSE
       "DB1146_PromptFree".ST01.Z05RetIng := FALSE;
   END_IF;
   // 含义：将 #ST01.Z05.ExtErr AND NOT ("ASMMode_M") 赋给 "DB1148_PromptBeeper".ST01.Z05ExtErr
   "DB1148_PromptBeeper".ST01.Z05ExtErr := #ST01.Z05.ExtErr AND NOT ("ASMMode_M");
   // 含义：将 #ST01.Z05.RetErr AND NOT ("ASMMode_M") 赋给 "DB1148_PromptBeeper".ST01.Z05RetErr
   "DB1148_PromptBeeper".ST01.Z05RetErr := #ST01.Z05.RetErr AND NOT ("ASMMode_M");
   // 含义：将 (#ST01.Z05.ExtEVT AND NOT ("ASMMode_M")) OR (#ST01.Z05.ExtEVT AND "AutoMode_M") 赋给 "DB1900_Communication_PC".Send.Z05Ext
   "DB1900_Communication_PC".Send.Z05Ext := (#ST01.Z05.ExtEVT AND NOT ("ASMMode_M")) OR (#ST01.Z05.ExtEVT AND "AutoMode_M");
   // 含义：将 (#ST01.Z05.RetEVT AND NOT ("ASMMode_M")) OR (#ST01.Z05.RetEVT AND "AutoMode_M") 赋给 "DB1900_Communication_PC".Send.Z05Ret
   "DB1900_Communication_PC".Send.Z05Ret := (#ST01.Z05.RetEVT AND NOT ("ASMMode_M")) OR (#ST01.Z05.RetEVT AND "AutoMode_M");
   // 含义：条件 "IToolAtPos" AND "DB1900_Communication_PC".Recv.Z05ExtTPPB 成立时，将 FALSE 传送到 "QZ14ExtEvt"
   IF "IToolAtPos" AND "DB1900_Communication_PC".Recv.Z05ExtTPPB THEN
       "QZ14ExtEvt" := FALSE;
   END_IF;
   // 含义：条件 "IToolAtPos" AND "DB1900_Communication_PC".Recv.Z05ExtTPPB 成立时，将 TRUE 传送到 "QZ14RetEvt"
   IF "IToolAtPos" AND "DB1900_Communication_PC".Recv.Z05ExtTPPB THEN
       "QZ14RetEvt" := TRUE;
   END_IF;
   // 含义：将 (("IToolAtPos" AND "DB1900_Communication_PC".Recv.Z05ExtTPPB) AND ("DB1900_Communication_PC".Recv.Current_2 >= 0.5)) 赋给 "DB1900_Communication_PC".Send.ToolPowerOn
   "DB1900_Communication_PC".Send.ToolPowerOn := (("IToolAtPos" AND "DB1900_Communication_PC".Recv.Z05ExtTPPB) AND ("DB1900_Communication_PC".Recv.Current_2 >= 0.5));
   // 含义：将 "IToolAtPos" AND "DB1900_Communication_PC".Recv.Z05ExtTPPB 赋给 "QWaterContactor"
   "QWaterContactor" := "IToolAtPos" AND "DB1900_Communication_PC".Recv.Z05ExtTPPB;
   // 含义：条件 "IToolAtPos" AND "DB1900_Communication_PC".Recv.Z05RetTPPB 成立时，将 TRUE 传送到 "QZ14ExtEvt"
   IF "IToolAtPos" AND "DB1900_Communication_PC".Recv.Z05RetTPPB THEN
       "QZ14ExtEvt" := TRUE;
   END_IF;
   // 含义：条件 "IToolAtPos" AND "DB1900_Communication_PC".Recv.Z05RetTPPB 成立时，将 FALSE 传送到 "QZ14RetEvt"
   IF "IToolAtPos" AND "DB1900_Communication_PC".Recv.Z05RetTPPB THEN
       "QZ14RetEvt" := FALSE;
   END_IF;
   // 含义：条件 NOT ("IToolAtPos") 成立时，将 FALSE 传送到 "QZ14ExtEvt"
   IF NOT ("IToolAtPos") THEN
       "QZ14ExtEvt" := FALSE;
   END_IF;
   // 含义：条件 NOT ("IToolAtPos") 成立时，将 FALSE 传送到 "QZ14RetEvt"
   IF NOT ("IToolAtPos") THEN
       "QZ14RetEvt" := FALSE;
   END_IF;

